(* IEC 61131-3 sources: daoli-st-library/DL_Process (part 31) *)

(* ---- FB_DL_EfEmoInterlock.st ---- *)
(*==============================================================================
 * 组件名称 (Component)  : FB_DL_EfEmoInterlock
 * 所属子库 (Sublibrary) : DL_Process
 * 当前版本 (Version)    : 1.0.0
 * 兼容性   (Platform)   : CODESYS 3.5+ / TwinCAT 3 / 汇川 InoProShop / 施耐德 Machine Expert
 *                         仅依赖 Standard.library（R_TRIG），零厂商私有库
 * 功能描述 (Function)   : EFEM 机械手互锁矩阵（域专用条件源）。
 *                         把 EFEM 域的四类条件源汇总成"机械手可否运动"的单一许可位，并追踪**首因**：
 *                           ① 门类（4 点）：安全门 / 维护门关到位，任一门未关 → 禁止运动；
 *                           ② 阀类（4 点）：隔离阀关到位，任一阀未关 → 禁止运动；
 *                           ③ 真空类（4 点）：吸盘/腔体真空建立，任一路失真空 → 禁止运动；
 *                           ④ 位置类（4 点）：机构在安全位，任一路越位 → 禁止运动。
 *                         判据顺序固定为"门 → 阀 → 真空 → 位置"（安全优先级由高到低），
 *                         首个失败项即首因；首因**锁存到全部条件恢复**才清零（不在故障期按当下输入
 *                         反复改写，R152/R190），HMI 因此能看到"是谁先拦的"。
 *                         验收向量：
 *                           ① 16 点全 TRUE → bMotionPermit = TRUE，eFirstCause = eNone
 *                           ② 门 3 未关 + 真空 1 失真空 → 首因 = eDoor，iFirstIdx = 3（门优先）
 *                           ③ 门恢复、真空 1 仍失 → 首因改判为 eVac，iFirstIdx = 1
 *                           ④ 三点同时失败 → 只报扫描序最靠前的一处（首因唯一）
 * 接口     (Interface)  : 入 abDoorClosed / abValveClosed / abVacOk / abInSafePos 四张 4 点条件表、
 *                         bMotionReq 运动请求（仅用于判定是否"曾经放行过"，不参与互锁本体）、
 *                         bReset 首因复位沿；
 *                         出 bMotionPermit 运动许可、bAnyBlocked 当前存在阻断、
 *                         eFirstCause 首因类别、iFirstIdx 首因点号（1..4，0 = 无）、
 *                         bFirstLatched 首因处于锁存态、eState 相、eCause 成因、bError 故障标志。
 * 边界     (Boundary)   : ① **属主边界（写死）：本件只做"EFEM 域条件源汇总与首因追踪"，
 *                         不内嵌通用互锁矩阵判据**（通用矩阵属 `FB_DL_InterlockMatrix`，
 *                         两件分工：本件是域条件源适配层，那件是任意规模矩阵求值器）；
 *                         本件也不驱动机械手运动、不做安全回路硬线判断（硬线由安全继电器负责）；
 *                         ② **数组边界**：四张表以字面量上界 4 声明（R104），扫描以常量
 *                         DL_EMI_N 之展开，不做动态下标，越界结构性不可能；
 *                         ③ **首因锁存解除式**：bReset 上升沿 ∨ 全部条件恢复（两式自证可满足：
 *                         前者为外部引脚恒可达，后者由条件源自身恢复触发）；
 *                         ④ **非门控输出**：eFirstCause 在锁存态下回放锁存值，不按当下输入重算（R152）；
 *                         ⑤ 零全局变量、零物理地址。
 * 分工声明 (Scope)      : 本件只管"EFEM 域四类条件源的首因判定"。不接管：门锁硬件状态诊断、
 *                         真空度模拟量判读、机械手轨迹安全校验（分别属门件/模拟量件/运动件）。
 * 来源标签 (Source Tag) : ROADMAP 空勾真缺口（EFEM 互锁，自研 clean-room）
 * 码表     (Codes)      : 本件不占用任何全局数字码位（零码位范式 R297）；诊断由 BOOL + ENUM 出口承担。
 * 红线自检 (Redline)    : R1 ✓ 零 GVL/VAR_EXTERNAL ｜ R2 ✓ 零 %I/%Q/%M ｜ R3 ✓ 纯 IEC 61131-3
 *                         R4 ✓ 定长展开无动态下标 + 首因唯一 + 解除式可满足 ｜ R5 ✓ 声明逐行同行双语注释
 *                         R6 ✓ ENUM+CASE 含 ELSE 兜底 ｜ R7 ✓ R_TRIG 段 0 无条件刷新（本件无 TON）
 * 修订历史 (Revision)   : 2026-11-19  v1.0.0  R47 首版（批次 3 · 序号 15）
 *==============================================================================*)

TYPE E_DL_EmiCause :
(
    eNone    := 0,   // 无阻断（全部条件满足） / No block, all conditions satisfied
    eDoor    := 1,   // 门未关到位（最高优先级） / Door not closed, highest priority
    eValve   := 2,   // 隔离阀未关到位 / Isolation valve not closed
    eVac     := 3,   // 真空失效 / Vacuum lost
    ePos     := 4,   // 机构不在安全位 / Mechanism off the safe position
    ePhaseBad:= 5    // 非法相位兜底 / Illegal phase fallback
);
END_TYPE

TYPE E_DL_EmiState :
(
    ePermit := 0,    // 放行相（条件全满足） / Permit, all conditions met
    eBlock  := 10,   // 阻断相（存在不满足条件） / Blocked
    eFault  := 90    // 故障相（内部非法，等复位） / Fault, awaiting reset
);
END_TYPE

FUNCTION_BLOCK FB_DL_EfEmoInterlock
VAR_INPUT
    abDoorClosed  : ARRAY[1..4] OF BOOL;   // 门关到位（1..4） [-] / Doors closed, points 1..4
    abValveClosed : ARRAY[1..4] OF BOOL;   // 隔离阀关到位（1..4） [-] / Valves closed, points 1..4
    abVacOk       : ARRAY[1..4] OF BOOL;   // 真空建立（1..4） [-] / Vacuum established, points 1..4
    abInSafePos   : ARRAY[1..4] OF BOOL;   // 机构在安全位（1..4） [-] / Mechanism in the safe position, points 1..4
    bMotionReq    : BOOL := FALSE;         // 机械手运动请求（诊断用，不参与互锁本体） [-] / Motion request, diagnostic only
    bReset        : BOOL := FALSE;         // 首因复位沿 [-] / First-cause reset edge
END_VAR
VAR_OUTPUT
    bMotionPermit : BOOL := FALSE;                      // 运动许可 [-] / Motion permit
    bAnyBlocked   : BOOL := FALSE;                      // 当前存在阻断（实时量） [-] / Any block present, live value
    eFirstCause   : E_DL_EmiCause := E_DL_EmiCause.eNone;   // 首因类别（锁存态回放） [-] / First cause, latched value
    iFirstIdx     : INT := 0;                           // 首因点号（1..4；0 = 无） [-] / First-cause point index, 0 = none
    bFirstLatched : BOOL := FALSE;                      // 首因处于锁存态 [-] / First cause currently latched
    eState        : E_DL_EmiState := E_DL_EmiState.ePermit; // 相出口 [-] / Phase outlet
    eCause        : E_DL_EmiCause := E_DL_EmiCause.eNone;   // 成因出口（与首因同源） [-] / Cause outlet
    bError        : BOOL := FALSE;                      // 故障标志（仅内部非法） [-] / Error flag
END_VAR
VAR
    _eState   : E_DL_EmiState := E_DL_EmiState.ePermit; // 内部相（CASE 唯一写入目标） / Internal phase
    _eCause   : E_DL_EmiCause := E_DL_EmiCause.eNone;  // 成因锁存量 / Latched cause
    _iIdx     : INT := 0;                               // 首因点号锁存量 / Latched first-cause index
    _bFault   : BOOL := FALSE;                          // 故障锁存位 / Latched fault bit
    _bBlocked : BOOL := FALSE;                          // 实时阻断量 / Live blocked flag
    _eNow     : E_DL_EmiCause := E_DL_EmiCause.eNone;  // 当拍首因（未锁存） / Live first cause
    _iNow     : INT := 0;                               // 当拍首因点号 / Live first-cause index
    rtReset   : R_TRIG;                                 // 复位沿实例，段 0 无条件调用 / Reset edge instance
END_VAR
VAR CONSTANT
    DL_EMI_N : INT := 4;              // 条件源点数（与四张表字面量上界同源，改动须同步） [点] / Points per source table
END_VAR

(* —— 段 0：沿实例无条件周期刷新（R228A；本件无 TON） —— *)
rtReset(CLK := bReset);                                  // 复位沿 / Reset edge

(* —— 段 1：单拍量预清零（锁存量 _eCause/_iIdx/_bFault 不入清单，R107） —— *)
bError      := FALSE;                                    // 故障标志预清（R45 配对） / Error preset
_bBlocked   := FALSE;                                    // 实时阻断量预清 / Live blocked preset
_eNow       := E_DL_EmiCause.eNone;                      // 当拍首因预置 / Live cause preset
_iNow       := 0;                                        // 当拍点号预置 / Live index preset

(* —— 段 2：首因扫描（定长展开，门 → 阀 → 真空 → 位置，安全优先级由高到低） —— *)
IF NOT abDoorClosed[1] THEN
    _eNow := E_DL_EmiCause.eDoor;  _iNow := 1;
ELSIF NOT abDoorClosed[2] THEN
    _eNow := E_DL_EmiCause.eDoor;  _iNow := 2;
ELSIF NOT abDoorClosed[3] THEN
    _eNow := E_DL_EmiCause.eDoor;  _iNow := 3;
ELSIF NOT abDoorClosed[4] THEN
    _eNow := E_DL_EmiCause.eDoor;  _iNow := 4;
ELSIF NOT abValveClosed[1] THEN
    _eNow := E_DL_EmiCause.eValve; _iNow := 1;
ELSIF NOT abValveClosed[2] THEN
    _eNow := E_DL_EmiCause.eValve; _iNow := 2;
ELSIF NOT abValveClosed[3] THEN
    _eNow := E_DL_EmiCause.eValve; _iNow := 3;
ELSIF NOT abValveClosed[4] THEN
    _eNow := E_DL_EmiCause.eValve; _iNow := 4;
ELSIF NOT abVacOk[1] THEN
    _eNow := E_DL_EmiCause.eVac;   _iNow := 1;
ELSIF NOT abVacOk[2] THEN
    _eNow := E_DL_EmiCause.eVac;   _iNow := 2;
ELSIF NOT abVacOk[3] THEN
    _eNow := E_DL_EmiCause.eVac;   _iNow := 3;
ELSIF NOT abVacOk[4] THEN
    _eNow := E_DL_EmiCause.eVac;   _iNow := 4;
ELSIF NOT abInSafePos[1] THEN
    _eNow := E_DL_EmiCause.ePos;   _iNow := 1;
ELSIF NOT abInSafePos[2] THEN
    _eNow := E_DL_EmiCause.ePos;   _iNow := 2;
ELSIF NOT abInSafePos[3] THEN
    _eNow := E_DL_EmiCause.ePos;   _iNow := 3;
ELSIF NOT abInSafePos[4] THEN
    _eNow := E_DL_EmiCause.ePos;   _iNow := 4;
ELSE
    _eNow := E_DL_EmiCause.eNone;  _iNow := 0;           // 全部满足：无首因 / All satisfied: no cause
END_IF
_bBlocked := (_eNow <> E_DL_EmiCause.eNone);             // 实时阻断量 / Live blocked flag

(* —— 段 3：首因锁存与解除（锁存期不按当下输入重算，R152） —— *)
IF _bBlocked THEN
    IF (_eCause = E_DL_EmiCause.eNone) THEN
        _eCause := _eNow;                                // 首次出现阻断：记首因 / First block: latch the cause
        _iIdx   := _iNow;                                // 记首因点号 / Latch the point
    END_IF
ELSE
    _eCause := E_DL_EmiCause.eNone;                      // 全部恢复：首因自动解除（解除式路径 1） / All clear: auto-release
    _iIdx   := 0;
END_IF
IF rtReset.Q THEN
    _eCause := E_DL_EmiCause.eNone;                      // 人工复位：清首因（解除式路径 2，恒可达） / Manual reset
    _iIdx   := 0;
    _bFault := FALSE;                                    // 同时清内部故障锁存 / Clear the internal fault latch
END_IF

(* —— 段 4：相迁移（许可 / 阻断两相；非法兜底） —— *)
CASE _eState OF

E_DL_EmiState.ePermit:
    IF _bBlocked THEN
        _eState := E_DL_EmiState.eBlock;                 // 出现阻断：进阻断相 / Enter the blocked phase
    END_IF

E_DL_EmiState.eBlock:
    IF NOT _bBlocked THEN
        _eState := E_DL_EmiState.ePermit;                // 条件恢复：回放行相 / Conditions recovered
    END_IF

E_DL_EmiState.eFault:
    ;                                                    // 故障相：由段 3 复位沿迁出 / Exit via the reset edge

ELSE
    _eCause := E_DL_EmiCause.ePhaseBad;                  // 归因：非法相位 / Cause: illegal phase
    _bFault := TRUE;                                     // 锁存 / Latch
    _eState := E_DL_EmiState.eFault;                     // 强拉故障相 / Force fault phase

END_CASE

(* —— 段 5：出口单点映射（许可位与本拍阻断量同源；首因回放锁存值，R191） —— *)
bMotionPermit := (NOT _bBlocked) AND (NOT _bFault) AND (_eState = E_DL_EmiState.ePermit);   // 运动许可 / Motion permit
bAnyBlocked   := _bBlocked;                                                                  // 实时阻断出口 / Live blocked outlet
eFirstCause   := _eCause;                                                                    // 首因出口（锁存回放） / First-cause outlet
iFirstIdx     := _iIdx;                                                                      // 首因点号出口 / First-cause index outlet
bFirstLatched := (_eCause <> E_DL_EmiCause.eNone);                                            // 首因锁存态出口 / Latched flag outlet
eState        := _eState;                                                                    // 相出口 / Phase outlet
eCause        := _eCause;                                                                    // 成因出口 / Cause outlet
bError        := _bFault OR (_bBlocked AND _bFault);                                          // 故障标志（仅内部非法） / Error flag

END_FUNCTION_BLOCK

(* ---- FB_DL_ElectrodeGapMark.st ---- *)
(*==============================================================================
 * 组件名称 (Component)  : FB_DL_ElectrodeGapMark
 * 所属子库 (Sublibrary) : DL_Process
 * 当前版本 (Version)    : 1.0.0
 * 兼容性 (Platform)     : CODESYS 3.5+ / TwinCAT 3 / 汇川 InoProShop / 施耐德 Machine Expert
 *                         仅依赖 Standard.library（R_TRIG / ABS），零厂商私有库
 * 功能描述 (Function)   : 极片留白区（Gap）位置标记与对齐判定。视觉/传感器
 *                         以 WORD 位域（每扇区 1 位）给出 Gap 标志，本件在
 *                         同步沿锁存编码位置为留白标记点，与上一标记点间距
 *                         对比组态节距判对齐（偏差超容差即 bAlignBad），并
 *                         统计位域有效位数。与 ScreenPrintAlign（丝印对位）
 *                         分工：本件面向极片 Gap 位域提取 + 留白带节距判定。
 * 来源标签 (Origin)     : ROADMAP §13.x P1（L626），自研 clean-room
 * 边界语义 (Boundary)   : ① 节距 <= eps 或容差 <= 0 → 组态故障锁存；
 *                         ② 位置 NaN 拍拒收标记（不锁存不判对齐）；
 *                         ③ 首个标记点（无前点）只锁存不判对齐（bAlignOk 缺省
 *                         FALSE，判定自第二个标记点起）；
 *                         ④ 位域统计移位量 0..15 结构性 < 16 位宽（R48 安全）。
 * 输出语义 (Fallback)   : 【R191】bEnable = FALSE → 标记/判定输出保持末值
 *                         （标记是资产属性不随失能消失）；eFault 相 → 冻结
 *                         + bError = TRUE。
 * 码位     (Codes)      : 按 R297 范式零 16# 码位硬编码；错误出口 BOOL+ENUM(eCause)。
 * 红线自检 (Redline)    : 7 项红线已自检：R1 零全局 ✓｜R2 零物理地址 ✓｜R3 纯 IEC ✓
 *                         R4 除零（节距 eps 闸）/NaN 拒收/组态闸 ✓
 *                         R5 双语同行注释 ✓｜R6 CASE 带 ELSE 兜底迁 eFault ✓
 *                         R7 R_TRIG 段 0 无条件刷新 ✓
 * 验收向量 (Acceptance) : V1 节距 100、容差 2：标记点 1000 → 1101（差 101）
 *                         → bAlignOk=TRUE，fDev=1.0；
 *                         V2 标记点 1000 → 1090（差 90，偏差 -10 超容差）
 *                         → bAlignOk=FALSE，bAlignBad=TRUE；
 *                         V3 uGapField=16#00F0 → nGapCnt=4。
 * 修订历史 (Revision)   : 2026-11-20  v1.0.0  R51 首版（批 1 · 序号 2）
 *==============================================================================*)
TYPE E_DL_EgmState :
(
    eIdle  := 0,                             (* 待使能 / Idle *)
    eTrack := 10,                            (* 标记跟踪运行 / Mark tracking *)
    eFault := 90                             (* 故障锁存相 / Fault latched phase *)
);
END_TYPE

TYPE E_DL_EgmCause :
(
    eNone       := 0,                        (* 无故障成因 / No cause *)
    eCfgIllegal := 1,                        (* 组态非法：节距/容差越域 / Illegal config *)
    ePhaseBad   := 2                         (* 非法相位兜底 / Illegal phase fallback *)
);
END_TYPE

FUNCTION_BLOCK FB_DL_ElectrodeGapMark
VAR_INPUT
    uGapField : WORD := 16#0000;             (* Gap 位域输入（每扇区 1 位，视觉给出）[-] / Gap bit field *)
    fPosNow   : LREAL := 0.0;                (* 当前编码位置 [mm] / Current encoder position *)
    fGapPitch : LREAL := 100.0;              (* 留白区节距，域 > eps [mm] / Gap pitch *)
    fTol      : LREAL := 2.0;                (* 节距对齐容差，域 > 0 [mm] / Pitch tolerance *)
    bSync     : BOOL := FALSE;               (* 视觉同步电平（上升沿锁标记点）[-] / Vision sync level *)
    bEnable   : BOOL := TRUE;                (* 使能 [-] / Enable *)
    bReset    : BOOL := FALSE;               (* 复位命令，上升沿清全部 [-] / Reset command *)
END_VAR
VAR_OUTPUT
    fMarkPos  : LREAL;                       (* 最新留白标记点位置 [mm] / Latest mark position *)
    fDev      : LREAL;                       (* 本标记点节距偏差（实测间距 - 节距）[mm] / Pitch deviation *)
    bAlignOk  : BOOL;                        (* 对齐判定（自第 2 个标记点起有效）[-] / Align verdict *)
    bAlignBad : BOOL;                        (* 对齐超差锁存（复位沿清）[-] / Align-fail latch *)
    nGapCnt   : INT;                         (* 位域有效位数 0..16 [位] / Set-bit count *)
    nMarkCnt  : UDINT;                       (* 累计标记点数 [点] / Total mark count *)
    eState    : E_DL_EgmState;               (* 状态出口 / State outlet *)
    eCause    : E_DL_EgmCause;               (* 故障成因出口 / Fault cause outlet *)
    bError    : BOOL;                        (* 故障锁存标志 [-] / Fault latch flag *)
END_VAR
VAR
    _eState  : E_DL_EgmState := E_DL_EgmState.eIdle;      (* 内部相位（CASE 唯一写入目标） / Internal phase *)
    _eCause  : E_DL_EgmCause := E_DL_EgmCause.eNone;      (* 故障成因锁存量 / Latched cause *)
    rtSync   : R_TRIG;                       (* 同步沿实例，段 0 无条件调用 / Sync edge instance *)
    rtReset  : R_TRIG;                       (* 复位沿实例，段 0 无条件调用 / Reset edge instance *)
    _fPrevMark : LREAL;                      (* 上一标记点位置 [mm] / Previous mark position *)
    _bHasPrev  : BOOL;                       (* 已有前点标志 [-] / Has previous mark *)
    _nCnt    : INT;                          (* 位域计数工作量 [-] / Bit count work *)
    _i       : INT;                          (* 位扫描游标（每趟重置，R227）[-] / Bit cursor *)
    _wMask   : WORD;                         (* 位掩码工作量 [-] / Bit mask work *)
    _nMark   : UDINT;                        (* 累计标记点数锁存 [点] / Mark count latch *)
    _fDev    : LREAL;                        (* 节距偏差派生量 [mm] / Deviation derived *)
    _bPosBad : BOOL;                         (* 位置非有限当拍量 [-] / Non-finite position *)
    _bFault  : BOOL;                         (* 故障锁存位 / Latched fault bit *)
    _bCfgBad : BOOL;                         (* 组态非法当拍量 / Illegal config this scan *)
END_VAR
VAR CONSTANT
    DL_EGM_EPS : LREAL := 1.0E-9;            (* 节距判零容差 [mm] / Pitch epsilon *)
END_VAR

(* —— 段 0：当拍判据派生 + 沿实例无条件刷新（R228A） —— *)
_bCfgBad := (fGapPitch <= DL_EGM_EPS) OR (fTol <= 0.0);   (* 组态闸（R151 全引脚） / Config gate *)
rtSync(CLK := bSync);                        (* 同步沿每拍必调 / Sync edge every scan *)
rtReset(CLK := bReset);                      (* 复位沿每拍必调 / Reset edge every scan *)
_bPosBad := (fPosNow <> fPosNow) OR ((fPosNow - fPosNow) <> (fPosNow - fPosNow));   (* 位置 NaN 自反 + Inf 差判 / Non-finite position *)

(* —— 段 1：单拍量预清零（R107） —— *)
_nCnt := 0;                                  (* 位计数预清（每趟重算，R285） / Bit count preset *)
_fDev := 0.0;                                (* 偏差预清 / Deviation preset *)
bAlignOk := FALSE;                           (* 对齐判定预清（判定拍内赋值，全路径覆盖） / Align preset *)

(* —— 段 2：复位沿处理（作用域：清故障 + 清标记点 + 清对齐锁存 + 清计数 + 迁 eIdle，R283 逐项声明） —— *)
IF rtReset.Q THEN
    _bFault := FALSE;                        (* 清故障锁存 / Clear fault *)
    _eCause := E_DL_EgmCause.eNone;          (* 清成因 / Clear cause *)
    _fPrevMark := 0.0;                       (* 清前点 / Clear previous mark *)
    _bHasPrev := FALSE;                      (* 清前点标志 / Clear has-prev *)
    bAlignBad := FALSE;                      (* 清超差锁存 / Clear fail latch *)
    fMarkPos := 0.0;                         (* 清标记出口 / Clear mark outlet *)
    fDev := 0.0;                             (* 清偏差出口 / Clear dev outlet *)
    _nMark := 0;                             (* 清累计计数 / Clear mark count *)
    _eState := E_DL_EgmState.eIdle;          (* 迁待机相 / Back to idle *)
END_IF

(* —— 段 3：组态闸故障锁存（R45 配对；锁存至复位沿，R189） —— *)
IF _bCfgBad AND NOT _bFault THEN
    _bFault := TRUE;                         (* 锁存故障位 / Latch fault *)
    _eCause := E_DL_EgmCause.eCfgIllegal;    (* 成因：组态非法 / Cause: illegal config *)
    _eState := E_DL_EgmState.eFault;         (* 同步迁故障相 / Migrate to fault *)
END_IF

(* —— 段 4：CASE 主状态机（ELSE 兜底迁 eFault，红线 6） —— *)
CASE _eState OF
    E_DL_EgmState.eIdle:                     (* 待机相 / Idle *)
        IF bEnable AND NOT _bFault THEN
            _eState := E_DL_EgmState.eTrack; (* 进入跟踪 / Enter track *)
        END_IF
    E_DL_EgmState.eTrack:                    (* 跟踪相：位域统计 + 同步沿标记判定 / Track *)
        IF NOT bEnable THEN
            _eState := E_DL_EgmState.eIdle;  (* 失能回待机 / Back to idle *)
        ELSE
            _i := 0;                         (* 位游标重置（R227） / Bit cursor reset *)
            _wMask := 16#0001;               (* 掩码起点（位 0） / Mask start *)
            WHILE _i <= 15 DO                (* 逐位统计（移位量 0..15 < 16 位宽，R48 安全） / Per-bit count *)
                IF (uGapField AND _wMask) <> 16#0000 THEN
                    _nCnt := _nCnt + 1;      (* 有效位计数 / Count set bit *)
                END_IF
                _wMask := SHL(_wMask, 1);    (* 掩码左移 1 位（常量移位量，R48） / Shift mask *)
                _i := _i + 1;                (* 游标递进 / Cursor advance *)
            END_WHILE
            IF rtSync.Q AND (NOT _bPosBad) THEN   (* 同步沿 + 位置有限：锁标记点 / Sync edge with finite pos *)
                IF _bHasPrev THEN
                    _fDev := (fPosNow - _fPrevMark) - fGapPitch;   (* 节距偏差派生（除法无涉，无除零） / Pitch deviation *)
                    bAlignOk := ABS(_fDev) <= fTol;   (* 对齐判定（容差闸） / Align verdict *)
                    IF NOT bAlignOk THEN
                        bAlignBad := TRUE;   (* 超差锁存至复位沿 / Latch align fail *)
                    END_IF
                    fDev := _fDev;           (* 偏差出口刷新 / Dev outlet *)
                END_IF
                _fPrevMark := fPosNow;       (* 前点更新 / Update previous *)
                fMarkPos := fPosNow;         (* 标记出口刷新 / Mark outlet *)
                _bHasPrev := TRUE;           (* 置前点标志 / Set has-prev *)
                _nMark := _nMark + 1;        (* 累计计数（UDINT 自然回绕可接受：17 亿标记点） / Count marks *)
            END_IF                           (* 位置坏值拍：不锁存不判定（边界②） / Bad pos: skip *)
        END_IF
    E_DL_EgmState.eFault:                    (* 故障相：冻结保持，仅复位沿出 / Fault *)
        ;                                    (* 锁存回放（R28） / Replay from latch *)
    ELSE                                     (* 非法相位兜底迁安全态 / Illegal phase fallback *)
        _eState := E_DL_EgmState.eFault;     (* 迁故障相 / To fault *)
        _bFault := TRUE;                     (* 同步锁存 / Latch *)
        _eCause := E_DL_EgmCause.ePhaseBad;  (* 成因：非法相位 / Cause: illegal phase *)
END_CASE

(* —— 段 5：出口映射（bError/eState 同源，R191） —— *)
nGapCnt := _nCnt;                            (* 位计数出口 / Bit count outlet *)
nMarkCnt := _nMark;                          (* 累计计数出口 / Mark count outlet *)
bError := _bFault;                           (* 故障标志镜像 / Fault flag mirror *)
eState := _eState;                           (* 状态出口 / State outlet *)
eCause := _eCause;                           (* 成因出口 / Cause outlet *)
END_FUNCTION_BLOCK

(* ---- FB_DL_ElectrolessBathReplenishCtrl.st ---- *)
(*
  DL Factory R83 | FB_DL_ElectrolessBathReplenishCtrl
  功能：按受镀面积与沉积速率算金属消耗，折算补加液量并做三态补加泵时序。
  开源溯源：无（clean-room 自研，依据公开工艺公式，来源=行业通用公式，许可证=MIT，借鉴点=公式结构）
  规则：R1-R21 全遵守
*)
TYPE E_DL_BathSt : ( eBathIdle := 0, eBathDose := 1, eBathFault := 2 ); END_TYPE // 补加三态枚举
FUNCTION_BLOCK FB_DL_ElectrolessBathReplenishCtrl
VAR_INPUT
    fLoadDm2    : REAL; // 在线受镀面积 [dm²] / In-line plated area [dm^2]
    fRateUmH    : REAL; // 沉积速率 [µm/h] / Deposition rate [um/h]
    fConcGpl    : REAL; // 槽液金属浓度 [g/L] / Bath metal concentration [g/L]
    fSpGpl      : REAL; // 目标维持浓度 [g/L] / Target maintained concentration [g/L]
    fAddConcGpl : REAL; // 补加液金属浓度 [g/L] / Replenisher metal concentration [g/L]
    bEnable     : BOOL; // 补加使能 / Dosing enable
    bReset      : BOOL; // 复位：清锁存码并回空闲相 / Reset: clear latched code, back to idle
END_VAR
VAR_OUTPUT
    fMetalGph : REAL; // 金属消耗速率 [g/h] / Metal consumption rate [g/h]
    fAddLph   : REAL; // 补加液流量指令 [L/h] / Replenisher flow command [L/h]
    xPump     : BOOL; // 补加泵运行输出 / Replenisher pump output
    iErrCode  : INT;  // 错误码，0=无错 / Error code, 0 = no error
END_VAR
VAR
    _eState : E_DL_BathSt := eBathIdle; // 当前状态，枚举初值一律 := / Current state, enum init with :=
    _iLatch : INT;        // 故障码锁存，仅 bReset 沿清除 / Latched fault code, reset edge only
    cNiGcm3 : REAL := 8.90; // 镍密度常量 [g/cm³]，已引用（R19）/ Nickel density [g/cm^3]
END_VAR
fMetalGph := 0.0; fAddLph := 0.0; xPump := FALSE;    // 出口预置：泵停（故障安全侧）
IF bReset THEN _iLatch := 0; iErrCode := 0; _eState := eBathIdle; END_IF  // 唯一清除边（R188）
// 非有限拦截 + 量纲自检 + 补加液浓度次序闸（R20/R21）
IF NOT (fLoadDm2 > -1.0E30 AND fLoadDm2 < 1.0E30) OR NOT (fRateUmH > -1.0E30 AND fRateUmH < 1.0E30) OR NOT (fConcGpl > -1.0E30 AND fConcGpl < 1.0E30) OR NOT (fSpGpl > -1.0E30 AND fSpGpl < 1.0E30) OR NOT (fAddConcGpl > -1.0E30 AND fAddConcGpl < 1.0E30) OR fLoadDm2 < 0.0 OR fRateUmH < 0.0 OR fSpGpl <= 0.0 OR fAddConcGpl <= fSpGpl THEN
    _eState := eBathFault; _iLatch := 9201; iErrCode := _iLatch; RETURN; // 故障拍不开泵
END_IF
// 金属消耗：1 dm² = 100 cm²、1 µm = 1E-4 cm，故每 dm²·µm = 0.01 cm³；乘 ρ 得 g
fMetalGph := fLoadDm2 * fRateUmH * 0.01 * cNiGcm3;   // 金属消耗速率 [g/h] / Metal consumption [g/h]
// 补加流量：g/h ÷ (补加浓度 - 维持浓度)[g/L] = L/h，浓度差分母显式零闸（R4/R21）
IF (fAddConcGpl - fSpGpl) > 1.0E-9 THEN fAddLph := fMetalGph / (fAddConcGpl - fSpGpl); ELSE fAddLph := 0.0; END_IF
CASE _eState OF  // 三态机：浓度偏低进补加相；退出两条（失去使能 / 浓度达标）
eBathIdle:
    IF bEnable AND fConcGpl < fSpGpl THEN _eState := eBathDose; END_IF  // 浓度偏低进补加 / Low conc, dose
eBathDose:
    xPump := TRUE;                                    // 补加相开泵 / Pump on in dose state
    IF NOT bEnable OR fConcGpl >= fSpGpl THEN _eState := eBathIdle; END_IF // 退出两条合并判 / Either exit
eBathFault:
    xPump := FALSE; iErrCode := _iLatch;              // 故障相停泵，故障码锁存回放 / Latched replay
ELSE
    _eState := eBathFault; _iLatch := 9203;           // 非法状态兜底拦截（R6）/ Illegal state fallback
END_CASE
END_FUNCTION_BLOCK

(* ---- FB_DL_ElectrolyteDosingSeq.st ---- *)
//==============================================================================
// 功能块：FB_DL_ElectrolyteDosingSeq ｜ 中文名称：电解液定量注液顺控（复杂度 H）
// 所属子库：DL_Process ｜ 版本：v1.0.1 ｜ 兼容：CODESYS V3.5+ / TwinCAT 3 / 汇川 InoProShop
// 功能描述：电解液定量注液节拍链——抽液 → 称重核对 → 粗注 → 细注 →
//           静置 → 完成，粗/细切换点按目标量占比驱动，秤读数全程监视
//           （回退判秤异常），中止走两段化（断输出使能 → 惰转窗 → 关阀）。
// 开源溯源 (Origin)：道莅原创实现（参考 ISA-88 相-步骤语义与注液机工程惯例 分类与参数域）
// 单位表：m[g] / 占比[倍] / 时间[ms] / 计数[次]
// 错误码表：16#0005_01E2 信息级（粗细切换点已达，不置 bError）/
//           16#0005_01E3 预留禁用（不得挪用）/ 16#0005_0318 故障级（目标
//           注液量 <= 0 或切换占比域外或确认窗组态越界（tSettleTime 为 0
//           或大于步 1 超时、xCoastAbort 时 tCoastTime <= 0），组态非法，
//           置 bError）/ 16#0005_0319
//           故障级（称重回退判秤异常，暂停顺控保持输出，置 bError）/
//           16#0005_031A 故障级兜底（状态机落 ELSE 或步超时，R90 复用，
//           置 bError 并全输出断）
// 状态机：E_DL_ElyteDosingPhase（八态：eIdle=0 / eVacuumDraw=10 /
//           eWeighCheck=20 / eCoarseFill=30 / eFineFill=40 / eSettle=50 /
//           eDone=60 / eFault=99）。【命名留档】派单枚举名 E_DL_DosingPhase
//           已被 FB_DL_BatchDosingControl 占用且成员不兼容，按 R70 唯一
//           属主纪律改用 E_DL_ElyteDosingPhase，全库唯一定义。中止两段化
//           不占相位（八态契约锁定），由 _uAbortStage 内部标志驱动。
// 边界行为：① fTargetMassG <= 0 或切换占比域外或确认窗/惰转窗组态越界
//           （tSettleTime 为 0 或 > 步 1 超时 DL_DOS_TO_WEIGH——否则步 1
//           稳定窗结构性超时；xCoastAbort 时 tCoastTime <= 0——否则中止段
//           A 永不收口）→ 故障 0318；② 称重回退
//           （fScaleMassG 比上拍小超容差，注液执行期）→ 故障 0319，暂停
//           顺控保持输出，bReset 清锁存；③ bAbort 两段化照 §4 修复件样板：
//           泵输出使能立即断、注液阀保持不动 → 惰转窗满 → 关阀，禁单拍
//           先停后关，机检断言：abort 拍不得出现关阀输出置位；④ 八态
//           CASE 每态显式 + ELSE 兜底 → 031A + 全输出断；⑤ 步超时（步进
//           器判超时）→ 031A 复用（R90，无专用码位）；⑥ 非有限秤读数归入
//           秤异常（0319 复用，R90）。
// 依赖纪律：Process → Level 0 组合调用合法——步进引擎组合调用
//           FB_DL_StepSequencer（DL_Base，接口已核实：bStart/abStepDone/
//           auStepTimeout/bAbort/bReset → nCurrentStep/bRunning/bDone/
//           bError/nFaultStep），步号映射表见下方注释；全库单调用点（每拍
 // *           恰好调用一次，防双调用边沿竞态）；防除零/防回绕/R79 防御齐备。
// 修订历史：v1.0.0 2026-11-17 首版（R23 派单 · ROADMAP 锂电 P1 §409 + ISA-88 相语义次源）
//           v1.0.1 2026-11-17 R23 终审修复：段 3 补组态一致性闸——tSettleTime
//           > 步 1 超时 T#5S 时稳定窗结构性超时（必报 031A 假故障）、
//           tCoastTime <= 0 时中止段 A 永不收口，均归入 0318 锁存，契约不变。
//==============================================================================

(*------------------------------------------------------------------------------
 * 枚举: E_DL_ElyteDosingPhase（归属本功能块，同文件发布，全库唯一定义）
 * 含义: 注液顺控相位，与步进器步号一一映射（见步号映射表）。
 *-----------------------------------------------------------------------------*)
TYPE E_DL_ElyteDosingPhase :
(
    eIdle       := 0,   // 空闲：等启动 / Idle, awaiting start
    eVacuumDraw := 10,  // 抽液：泵送电解液至计量腔（步 0） / Vacuum draw, pumping electrolyte, step 0
    eWeighCheck := 20,  // 称重核对：秤读数稳定窗（步 1） / Weigh check, scale stability window, step 1
    eCoarseFill := 30,  // 粗注：注液阀开，至粗细切换点（步 2） / Coarse fill to the switch point, step 2
    eFineFill   := 40,  // 细注：注液阀开，至目标量（步 3） / Fine fill to the target mass, step 3
    eSettle     := 50,  // 静置：浸润计时与终值复核（步 4） / Settling, soak window and final check, step 4
    eDone       := 60,  // 完成：放行，等启动撤销（步 5） / Done, released, step 5
    eFault      := 99   // 故障：组态/秤异常/步超时/非法状态 / Fault, config, scale, timeout or illegal state
);
END_TYPE

(*------------------------------------------------------------------------------
 * 步号映射表（步进器步号 → 相位枚举）：
 *   0 → eVacuumDraw ｜ 1 → eWeighCheck ｜ 2 → eCoarseFill ｜ 3 → eFineFill
 *   4 → eSettle ｜ 5 → eDone（步进器 bDone）｜ -1 → eIdle
 * 语义假设（头注释留档）：电子秤位于注液目标侧，注液过程中读数单调
 *   递增；已注量 = 读数 − 启动基线；抽液侧无秤反馈，以固定时长判完成。
 *-----------------------------------------------------------------------------*)
FUNCTION_BLOCK FB_DL_ElectrolyteDosingSeq
VAR_INPUT
    bStart        : BOOL;                   // 启动请求 [—]，上升沿生效 / Start request, rising edge
    bAbort        : BOOL;                   // 中止请求 [—]，任意拍生效 / Abort request, effective on any scan
    bReset        : BOOL;                   // 故障复位 [—]，上升沿清秤异常锁存 / Fault reset, rising edge clears the scale latch
    fTargetMassG  : LREAL;                  // 目标注液量 [克]，须 > 0 / Target dosing mass [g], must be > 0
    fCoarseFineKg : LREAL := 0.95;          // 粗/细切换点占目标比 [倍]，有效域 0..1 / Coarse-to-fine switch ratio [ratio], 0..1
    fScaleMassG   : LREAL;                  // 电子秤实时读数 [克]，注液目标侧质量 / Scale reading [g], target-side mass
    tSettleTime   : TIME  := T#2S;          // 静置浸润计时 [ms]，兼作称重稳定窗 / Soak time [ms], also the weigh stability window
    xCoastAbort   : BOOL  := TRUE;          // TRUE = 中止走惰转两段化（推荐）/ FALSE = 单拍中止（不推荐：残压回流风险） / Coast-stop abort sequencing enabled
    tCoastTime    : TIME  := T#2S;          // 泵惰转时间 [ms]：断使能到关阀的物理时序分隔窗 / Pump coast-down time [ms]
END_VAR
VAR_OUTPUT
    ePhase        : E_DL_ElyteDosingPhase;  // 注液相位 [—] / Dosing phase
    fDosedMassG   : LREAL;                  // 已注量 [克] = 读数 − 基线 / Dosed mass [g] = reading minus baseline
    bDosingOut    : BOOL;                   // 注液阀输出 [—] / Dosing valve output
    bPumpOut      : BOOL;                   // 泵输出 [—] / Pump output
    eErr          : UDINT;                  // 错误码，0 = 无错 / Error code, 0 = no error
    bError        : BOOL;                   // 故障级标志，仅故障级错误置位 / Fault-class flag, set only on fault-level codes
    bValid        : BOOL;                   // 输出可用标志 / Outputs usable flag
END_VAR
VAR
    fbSeq         : FB_DL_StepSequencer;    // 步进引擎（Level 0 组合调用，单调用点） / Step engine, Level 0 composition, single call site
    fbDraw        : TON;                    // 抽液计时（步 0 完成判据），段 6 无条件刷新 [ms] / Draw timer, step 0 done criterion
    fbStable      : TON;                    // 称重稳定窗（步 1 完成判据），段 6 无条件刷新 [ms] / Weigh stability window, step 1 done criterion
    fbSettle      : TON;                    // 静置计时（步 4 完成判据），段 6 无条件刷新 [ms] / Settle timer, step 4 done criterion
    fbCoast       : TON;                    // 泵惰转计时（中止第一段），段 6 无条件刷新 [ms] / Pump coast timer, abort stage A
    _abStepDone   : ARRAY[0..15] OF BOOL;   // 步完成信号（本件按判据维护） / Step-done levels, maintained by this FB
    _auStepTimeout: ARRAY[0..15] OF TIME;   // 每步超时 [ms]，0 = 不监控 / Per-step timeout [ms], zero = not monitored
    _ePhase       : E_DL_ElyteDosingPhase := E_DL_ElyteDosingPhase.eIdle; // 当前相位 / Current phase
    _fBaseMassG   : LREAL;                  // 注液基线质量 [克]，启动拍锁定 / Baseline mass [g], locked at start
    _fScalePrevG  : LREAL;                  // 上拍秤读数快照 [克] / Previous-scan scale snapshot [g]
    _uAbortStage  : UINT;                   // 中止段号 [—]，0 = 无 / 1 = 惰转 / 2 = 已关阀 / Abort stage, zero none, one coast, two closed
    _bSeqStart    : BOOL;                   // 步进器启动沿请求（单调用点输入） / Sequencer start edge request
    _bStartPrev   : BOOL;                   // 启动命令上拍电平快照 / Previous-scan level of the start command
    _bInit        : BOOL := FALSE;          // 首扫标志，初值 FALSE 取非判定 / First-scan flag, tested negated
    _bParamBad    : BOOL;                   // 参数非法锁存 / Illegal parameter latch
    _bScaleErr    : BOOL;                   // 秤异常锁存（bReset 清除） / Scale fault latch, cleared by bReset
    _bIllegal     : BOOL;                   // 非法状态标志 / Illegal state flag
    _bInfoCoarse  : BOOL;                   // 粗细切换信息当拍标志 / Coarse switch info flag of this scan
END_VAR
VAR CONSTANT
    DL_DOS_TOL_G   : LREAL := 0.5;          // 秤稳定/回退容差 [克] / Scale stability and regression tolerance [g]
    DL_DOS_DRAW_T  : TIME  := T#5S;         // 抽液固定时长 [ms]，抽液无秤反馈侧判据的工程缺省 / Fixed draw duration [ms]
    DL_DOS_TO_DRAW : TIME  := T#8S;         // 步 0 超时 [ms] / Step 0 timeout [ms]
    DL_DOS_TO_WEIGH: TIME  := T#5S;         // 步 1 超时 [ms] / Step 1 timeout [ms]
    DL_DOS_TO_COARSE: TIME := T#60S;        // 步 2 超时 [ms] / Step 2 timeout [ms]
    DL_DOS_TO_FINE : TIME  := T#120S;       // 步 3 超时 [ms] / Step 3 timeout [ms]
    DL_DOS_TO_SETTLE: TIME := T#10S;        // 步 4 超时 [ms] / Step 4 timeout [ms]
    DL_DOS_INF     : LREAL := 1.7976931348623157E308; // LREAL 幅值上限 / LREAL magnitude ceiling
END_VAR

(*------------------------------------------------------------------------------
 * 段 1｜每拍预置：双输出先全断（安全侧），单拍标志预清零
 *      Both outputs cleared first, fail-safe, one-shot flags pre-cleared
 *-----------------------------------------------------------------------------*)
bDosingOut  := FALSE;                       // 注液阀输出先清（安全侧） / Dosing output cleared first
bPumpOut    := FALSE;                       // 泵输出先清（安全侧） / Pump output cleared first
fDosedMassG := 0.0;                         // 已注量每拍重算 / Dosed mass recomputed
eErr        := 16#0000_0000;                // 错误码每拍重算 / Error code recomputed
bError      := FALSE;                       // 故障标志每拍重算 / Fault flag recomputed
bValid      := FALSE;                       // 可用标志每拍重算 / Usable flag recomputed
_bIllegal   := FALSE;                       // 非法状态标志预清零 / Illegal flag pre-cleared
_bInfoCoarse := FALSE;                     // 粗细切换信息预清零 / Coarse info pre-cleared
_bSeqStart  := FALSE;                       // 步进器启动沿请求预清零 / Sequencer start request pre-cleared

(*------------------------------------------------------------------------------
 * 段 2｜首扫初始化：步超时表一次装配
 *      First-scan initialisation, the timeout table assembled once
 *-----------------------------------------------------------------------------*)
IF NOT _bInit THEN
    _ePhase := E_DL_ElyteDosingPhase.eIdle; // 相位空闲起步 / Phase starts idle
    _auStepTimeout[0] := DL_DOS_TO_DRAW;    // 步 0 抽液超时 / Step 0 draw timeout
    _auStepTimeout[1] := DL_DOS_TO_WEIGH;   // 步 1 称重超时 / Step 1 weigh timeout
    _auStepTimeout[2] := DL_DOS_TO_COARSE;  // 步 2 粗注超时 / Step 2 coarse timeout
    _auStepTimeout[3] := DL_DOS_TO_FINE;    // 步 3 细注超时 / Step 3 fine timeout
    _auStepTimeout[4] := DL_DOS_TO_SETTLE;  // 步 4 静置超时 / Step 4 settle timeout
    _auStepTimeout[5] := T#0MS;             // 步 5 完成态不监控 / Step 5 not monitored
    _fScalePrevG := 0.0;                    // 秤快照从零起步 / Scale snapshot starts at zero
    _uAbortStage := 0;                      // 中止段号从零起步 / Abort stage starts at zero
    _bInit := TRUE;                         // 首扫只做一次 / The first scan runs once
END_IF

(*------------------------------------------------------------------------------
 * 段 3｜参数与输入防御闸（R79 双侧幅值判 + 占比域闸）
 *      Parameter and input defense gates
 *-----------------------------------------------------------------------------*)
IF (fTargetMassG <> fTargetMassG) OR (ABS(fTargetMassG) > DL_DOS_INF) OR (fTargetMassG <= 0.0) THEN
    _bParamBad := TRUE;                     // 目标量非法锁存 / Illegal target latched
END_IF
IF (fScaleMassG <> fScaleMassG) OR (ABS(fScaleMassG) > DL_DOS_INF) THEN
    _bScaleErr := TRUE;                     // 秤读数非有限归入秤异常（0319 复用，R90） / Non-finite scale folded into the scale fault
END_IF
IF (fCoarseFineKg < 0.0) OR (fCoarseFineKg > 1.0) THEN
    _bParamBad := TRUE;                     // 切换占比域外锁存 / Switch ratio out of range latched
END_IF
IF (tSettleTime <= T#0MS) OR (tSettleTime > DL_DOS_TO_WEIGH) THEN
    _bParamBad := TRUE;                     // 确认窗组态越界：为 0 或大于步 1 超时（结构性超时）锁存 / Confirm window out of range, latched
END_IF
IF xCoastAbort AND (tCoastTime <= T#0MS) THEN
    _bParamBad := TRUE;                     // 惰转窗组态越界：两段化中止永不收口锁存 / Coast window out of range, latched
END_IF

(*------------------------------------------------------------------------------
 * 段 4｜称重回退检测（注液执行期）：比上拍小超容差 → 0319 锁存
 *      Scale regression detection during the dosing execution phases
 *-----------------------------------------------------------------------------*)
IF (_ePhase = E_DL_ElyteDosingPhase.eCoarseFill)
   OR (_ePhase = E_DL_ElyteDosingPhase.eFineFill)
   OR (_ePhase = E_DL_ElyteDosingPhase.eSettle) THEN
    IF fScaleMassG < (_fScalePrevG - DL_DOS_TOL_G) THEN
        _bScaleErr := TRUE;                 // 称重回退锁存（暂停顺控保持输出） / Scale regression latched, sequencing paused
    END_IF
END_IF
_fScalePrevG := fScaleMassG;                // 快照推进 / Snapshot advanced

(*------------------------------------------------------------------------------
 * 段 5｜中止入口（任意拍生效；中止族态内不重复触发）与复位
 *      Abort entry, effective on any scan, not re-triggered in the family
 *-----------------------------------------------------------------------------*)
IF bAbort AND (_uAbortStage = 0)
   AND (_ePhase = E_DL_ElyteDosingPhase.eVacuumDraw
        OR _ePhase = E_DL_ElyteDosingPhase.eWeighCheck
        OR _ePhase = E_DL_ElyteDosingPhase.eCoarseFill
        OR _ePhase = E_DL_ElyteDosingPhase.eFineFill
        OR _ePhase = E_DL_ElyteDosingPhase.eSettle) THEN
    _uAbortStage := 1;                      // 进中止段 A（惰转） / Enter abort stage A, coast
END_IF
IF _uAbortStage >= 1 THEN
    IF (NOT bStart) AND (_uAbortStage = 2) THEN
        _uAbortStage := 0;                  // 关阀已完成且启动撤销，回空闲 / Close done and start dropped, back to idle
        _ePhase      := E_DL_ElyteDosingPhase.eIdle; // 相位回空闲 / Phase back to idle
    END_IF
END_IF
IF bReset THEN
    _bScaleErr := FALSE;                    // 复位清秤异常锁存 / Reset clears the scale latch
END_IF

(*------------------------------------------------------------------------------
 * 段 6｜四只计时无条件刷新（R40：CASE 之外每拍必调，各司其职不复用）
 *      Four timers refreshed unconditionally per R40
 *-----------------------------------------------------------------------------*)
fbDraw(IN := (_ePhase = E_DL_ElyteDosingPhase.eVacuumDraw) AND (_uAbortStage = 0),
       PT := DL_DOS_DRAW_T);               // 抽液计时 / Draw timer
fbStable(IN := (_ePhase = E_DL_ElyteDosingPhase.eWeighCheck) AND (_uAbortStage = 0)
              AND (ABS(fScaleMassG - _fBaseMassG) < DL_DOS_TOL_G), PT := tSettleTime); // 称重稳定窗 / Weigh stability window
fbSettle(IN := (_ePhase = E_DL_ElyteDosingPhase.eSettle) AND (_uAbortStage = 0), PT := tSettleTime); // 静置计时 / Settle timer
fbCoast(IN := (_uAbortStage = 1), PT := tCoastTime); // 中止惰转计时（段 A） / Abort coast timer, stage A

(*------------------------------------------------------------------------------
 * 段 7｜步进器单调用点（每拍恰好一次）与步完成判据装配
 *      Single sequencer call site and the step-done criteria assembly
 *-----------------------------------------------------------------------------*)
_bSeqStart := bStart AND (NOT _bStartPrev) AND (_ePhase = E_DL_ElyteDosingPhase.eIdle)
              AND (NOT _bParamBad) AND (NOT _bScaleErr); // 启动沿（空闲且组态合法） / Start edge in idle with a legal configuration
_bStartPrev := bStart;                      // 电平快照推进 / Level snapshot advanced

IF (_ePhase <> E_DL_ElyteDosingPhase.eIdle) AND (_ePhase <> E_DL_ElyteDosingPhase.eFault)
   AND (_uAbortStage = 0) THEN
    _abStepDone[0] := fbDraw.Q;             // 步 0 完成：抽液计时满 / Step 0 done, draw elapsed
    _abStepDone[1] := fbStable.Q;           // 步 1 完成：秤读数稳定窗满 / Step 1 done, stability window elapsed
    _abStepDone[2] := (fScaleMassG - _fBaseMassG) >= (fTargetMassG * fCoarseFineKg); // 步 2 完成：达粗细切换点 / Step 2 done, switch point reached
    _abStepDone[3] := (fScaleMassG - _fBaseMassG) >= fTargetMassG; // 步 3 完成：达目标量 / Step 3 done, target reached
    _abStepDone[4] := fbSettle.Q;           // 步 4 完成：静置计时满 / Step 4 done, settle elapsed
    _abStepDone[5] := TRUE;                 // 步 5 完成态恒成 / Step 5 always done
    IF _abStepDone[2] AND (_ePhase = E_DL_ElyteDosingPhase.eCoarseFill) THEN
        _bInfoCoarse := TRUE;               // 粗细切换点已达（信息级） / Switch point reached, info
    END_IF
END_IF

fbSeq(bStart := _bSeqStart, abStepDone := _abStepDone, auStepTimeout := _auStepTimeout,
      bHold := FALSE, bSingleStep := FALSE, bAdvance := FALSE,
      bAbort := (_uAbortStage >= 1), bReset := FALSE); // 步进器唯一调用点 / The only sequencer call site

IF _uAbortStage = 1 THEN
    IF fbCoast.Q THEN
        _uAbortStage := 2;                  // 惰转窗满，进中止段 B（关阀） / Coast elapsed, abort stage B, close
    END_IF
END_IF

(*------------------------------------------------------------------------------
 * 段 8｜相位机（只做迁移与步进对账；输出在段 9 按相置位）
 *      Phase machine, transitions and step reconciliation only
 *-----------------------------------------------------------------------------*)
CASE _ePhase OF

    E_DL_ElyteDosingPhase.eIdle:           // 空闲：启动沿锁定基线进抽液
        IF _bSeqStart THEN
            _fBaseMassG := fScaleMassG;     // 基线锁定 / Baseline locked
            _ePhase     := E_DL_ElyteDosingPhase.eVacuumDraw; // 进抽液相 / To the draw phase
        END_IF

    E_DL_ElyteDosingPhase.eVacuumDraw:     // 抽液：步进器推进到步 1 即转称重
        IF fbSeq.bError THEN
            _ePhase := E_DL_ElyteDosingPhase.eFault; // 步超时，故障 / Step timeout, fault
        ELSIF (fbSeq.nCurrentStep = 1) THEN
            _ePhase := E_DL_ElyteDosingPhase.eWeighCheck; // 步进器已推进 / The sequencer advanced
        END_IF

    E_DL_ElyteDosingPhase.eWeighCheck:     // 称重核对：步进器推进到步 2 即转粗注
        IF fbSeq.bError THEN
            _ePhase := E_DL_ElyteDosingPhase.eFault; // 步超时，故障 / Step timeout, fault
        ELSIF (fbSeq.nCurrentStep = 2) THEN
            _ePhase := E_DL_ElyteDosingPhase.eCoarseFill; // 步进器已推进 / The sequencer advanced
        END_IF

    E_DL_ElyteDosingPhase.eCoarseFill:     // 粗注：步进器推进到步 3 即转细注
        IF fbSeq.bError THEN
            _ePhase := E_DL_ElyteDosingPhase.eFault; // 步超时，故障 / Step timeout, fault
        ELSIF (fbSeq.nCurrentStep = 3) THEN
            _ePhase := E_DL_ElyteDosingPhase.eFineFill; // 步进器已推进 / The sequencer advanced
        END_IF

    E_DL_ElyteDosingPhase.eFineFill:       // 细注：步进器推进到步 4 即转静置
        IF fbSeq.bError THEN
            _ePhase := E_DL_ElyteDosingPhase.eFault; // 步超时，故障 / Step timeout, fault
        ELSIF (fbSeq.nCurrentStep = 4) THEN
            _ePhase := E_DL_ElyteDosingPhase.eSettle; // 步进器已推进 / The sequencer advanced
        END_IF

    E_DL_ElyteDosingPhase.eSettle:         // 静置：步进器推进到步 5 即完成
        IF fbSeq.bError THEN
            _ePhase := E_DL_ElyteDosingPhase.eFault; // 步超时，故障 / Step timeout, fault
        ELSIF (fbSeq.nCurrentStep = 5) THEN
            _ePhase := E_DL_ElyteDosingPhase.eDone; // 步进器已推进 / The sequencer advanced
        END_IF

    E_DL_ElyteDosingPhase.eDone:           // 完成：等启动撤销回空闲
        IF NOT bStart THEN
            _ePhase := E_DL_ElyteDosingPhase.eIdle; // 回空闲 / Back to idle
        END_IF

    E_DL_ElyteDosingPhase.eFault:          // 故障：复位沿且原因消失回空闲
        IF bReset AND (NOT _bParamBad) AND (NOT _bScaleErr) THEN
            _ePhase := E_DL_ElyteDosingPhase.eIdle; // 回空闲 / Back to idle
        END_IF

    ELSE                                   // 非法状态兜底（R21：CASE 必带 ELSE）
        _bIllegal := TRUE;                 // 标记非法状态 / Flag the illegal state
        _ePhase   := E_DL_ElyteDosingPhase.eFault; // 回故障态（段 9 全断） / Back to fault, all outputs off
END_CASE

(*------------------------------------------------------------------------------
 * 段 9｜输出置位（次序即安全：泵先于阀；中止段 A 泵断使能、阀保持不动，
 *       机检断言：abort 拍不得出现关阀输出置位——段 A 阀输出 = 保持量）
 *      Output assignment, pump precedes the valve, abort stage A holds the valve
 *-----------------------------------------------------------------------------*)
CASE _ePhase OF
    E_DL_ElyteDosingPhase.eVacuumDraw:     // 抽液：泵运行 / Draw: pump runs
        bPumpOut := (_uAbortStage = 0);    // 中止段 A 泵使能立即断 / Pump enable cut immediately in abort stage A
    E_DL_ElyteDosingPhase.eCoarseFill:     // 粗注：阀开 / Coarse: valve open
        bDosingOut := (_uAbortStage = 0) OR (_uAbortStage = 1); // 段 A 阀保持，段 B 关阀 / Valve held in stage A, closed in stage B
    E_DL_ElyteDosingPhase.eFineFill:       // 细注：阀开 / Fine: valve open
        bDosingOut := (_uAbortStage = 0) OR (_uAbortStage = 1); // 段 A 阀保持，段 B 关阀 / Valve held in stage A, closed in stage B
    ELSE                                   // 其余相输出全断 / Otherwise all off
        bDosingOut := FALSE;               // 注液阀断 / Dosing off
        bPumpOut   := FALSE;               // 泵断 / Pump off
END_CASE
IF (NOT xCoastAbort) AND (_uAbortStage >= 1) THEN
    bDosingOut := FALSE;                   // 兼容路径：单拍中止（不推荐，残压回流风险） / Legacy single-scan abort, not recommended
    bPumpOut   := FALSE;                   // 泵同拍断 / Pump off the same scan
END_IF

fDosedMassG := fScaleMassG - _fBaseMassG;   // 已注量出口 [克] / Dosed mass outlet [g]
IF fDosedMassG < 0.0 THEN
    fDosedMassG := 0.0;                     // 负增量钳 0（换批/去皮期） / Negative delta clamped to zero
END_IF
ePhase := _ePhase;                          // 相位出口 / Phase outlet

IF _bIllegal THEN
    eErr   := 16#0005_031A;                 // 故障级：状态机兜底 / Fault: state machine fallback
    bError := TRUE;                         // 置故障标志 / Raise the fault flag
ELSIF _bParamBad THEN
    eErr   := 16#0005_0318;                 // 故障级：目标量或占比非法 / Fault: illegal target or ratio
    bError := TRUE;                         // 置故障标志 / Raise the fault flag
ELSIF _bScaleErr THEN
    eErr   := 16#0005_0319;                 // 故障级：称重回退判秤异常 / Fault: scale regression
    bError := TRUE;                         // 置故障标志 / Raise the fault flag
ELSIF fbSeq.bError THEN
    eErr   := 16#0005_031A;                 // 故障级：步超时复用兜底码（R90） / Fault: step timeout, code reused per R90
    bError := TRUE;                         // 置故障标志 / Raise the fault flag
ELSIF _bInfoCoarse THEN
    eErr := 16#0005_01E2;                   // 信息级：粗细切换点已达 / Info: switch point reached
END_IF

bValid := (NOT bError) AND (_ePhase <> E_DL_ElyteDosingPhase.eIdle); // 空闲/故障输出不可用 / Outputs unusable in idle or fault
END_FUNCTION_BLOCK

(* ---- FB_DL_ElectrolyteDosingTrend.st ---- *)
(*
  ==================================================================
  组件名 Component  : FB_DL_ElectrolyteDosingTrend
  分类   Category   : DL_Process
  版本   Version    : 1.0.0
  功能   Purpose    : 注液量趋势 SPG（统计过程判据）统计。逐次注液量进环窗，
                      窗满后给出均值、样本标准差、上下控制限（均值 ± k × 标准差）、
                      越限判据与连续同向趋势判据（连升 / 连降），并给目标带内
                      合格判据，用于注液泵磨损与堵塞的早期趋势预警。
  溯源   Origin     : 均值 / 标准差 / 控制限为公开统计过程控制口径；本件为 clean-room
                      实现，仅借鉴来源分类与参数域组织（来源标签 roadmap-p2-dosing），
                      道莅原创设计，未复制任何闭源代码行。
  平台   Platform   : 纯 IEC 61131-3（SQRT / REAL / R_TRIG，无私有库、无方言转换）
  作者   Author     : 道莅代码库 · PLC 编程专家（R55）
  ------------------------------------------------------------------
  边界 Boundary     :
                      一 本件只做统计与趋势判据，不调节注液泵、不改配方（属主边界）；
                      二 样本标准差按 n − 1 无偏口径，样本数小于 2 时不下结论；
                      三 方差由「平方和 − 和的平方 / n」推得，舍入致负值一律钳零（开方前闸）；
                      四 环窗遍历按时间序遍历，禁按数组下标序遍历（R194）；
                      五 无全局变量、无外部变量声明、无物理地址寻址。
  输出契约 Output contract:
                      fMeanMl / fStdMl / fUclMl / fLclMl 仅在样本数达标时更新，
                      否则保持上拍值；bOutOfCtrl 仅在最新样本越限时为真（单拍语义，
                      由调用方按需累计）；nTrendRun 正数为连升、负数为连降；
                      eCause 故障级成因与 bError 配对（R45），信息级永不置 bError。
  修订记录 Revision  :
    2026-11-20  v1.0.0  R55 首版（批 4 · 序号 15）
  ==================================================================
*)

TYPE E_DL_EdtTrend :
(
    eStable := 0,       // 平稳：最新与上一样本无明显方向 / stable, no clear direction between the last two samples
    eUp     := 10,      // 连升：连续同向上升 / rising, a run of increases
    eDown   := 20       // 连降：连续同向下降 / falling, a run of decreases
);
END_TYPE

TYPE E_DL_EdtCause :
(
    eNone       := 0,   // 无成因 / no cause
    eCfgIllegal := 1,   // 组态非法：窗口容量、系数或目标带越域（故障级，与 bError 配对）/ illegal config, window size, sigma factor or target band out of domain
    eNoSample   := 2,   // 样本数不足 2，统计量保持上拍值（信息级）/ fewer than two samples and the statistics hold, informational
    eBadSample  := 3    // 存在非有限样本，已拒收（信息级）/ non-finite samples were rejected, informational
);
END_TYPE

FUNCTION_BLOCK FB_DL_ElectrolyteDosingTrend
VAR_INPUT
    bEnable      : BOOL := TRUE;             // 使能，失能时不收样本 [-] / enable, no sample is accepted when disabled
    bReset       : BOOL := FALSE;           // 复位上升沿清故障锁存与全部统计 [-] / reset rising edge clears the fault latch and all statistics
    bSamplePulse : BOOL := FALSE;            // 单次注液量采样脉冲，上升沿收一条 [-] / single dose sample pulse, one sample per rising edge
    fVolMl       : REAL := 0.0;              // 本次注液量 [毫升] / dose volume of this shot [millilitre]
    fTargetMl    : REAL := 100.0;            // 目标注液量 [毫升]，域 大于零 / target dose volume [millilitre], domain above zero
    fTolPct      : REAL := 2.0;              // 目标带容差 [百分比]，域 大于零 / target band tolerance [percent], domain above zero
    nWinSize     : INT := 20;                // 统计窗样本数 [个]，域 2..64 / statistics window size [count], domain 2 to 64
    fSigmaK      : REAL := 3.0;              // 控制限系数（倍标准差）[倍]，域 1..6 / control limit factor in standard deviations [factor], domain 1 to 6
END_VAR
VAR_OUTPUT
    fMeanMl      : REAL := 0.0;              // 窗口均值 [毫升] / window mean [millilitre]
    fStdMl       : REAL := 0.0;              // 窗口样本标准差（n − 1 口径）[毫升] / window sample standard deviation over n minus one [millilitre]
    fUclMl       : REAL := 0.0;              // 上控制限 [毫升] / upper control limit [millilitre]
    fLclMl       : REAL := 0.0;              // 下控制限 [毫升]，可为负 / lower control limit, may be negative [millilitre]
    nSampleCnt   : INT := 0;                 // 窗口有效样本数 [个] / valid sample count in the window
    bOutOfCtrl   : BOOL := FALSE;            // 最新样本越控制限 [-] / the newest sample is beyond a control limit
    bHasStats    : BOOL := FALSE;            // 统计量是否已可交付 [-] / the statistics are deliverable
    bInTarget    : BOOL := FALSE;            // 最新样本落在目标带内 [-] / the newest sample is inside the target band
    nTrendRun    : INT := 0;                 // 连续同向计数（正连升 / 负连降）[次] / signed run length, positive rising and negative falling [count]
    eTrend       : E_DL_EdtTrend := E_DL_EdtTrend.eStable; // 趋势出口 [枚举] / trend outlet [enum]
    nRejectCnt   : INT := 0;                 // 累计拒收样本数（饱和到上限）[个] / total rejected samples, saturated [count]
    eCause       : E_DL_EdtCause := E_DL_EdtCause.eNone; // 成因出口 [枚举] / cause outlet [enum]
    bError       : BOOL := FALSE;            // 故障锁存标志 [-] / fault latch flag
END_VAR
VAR
    rtSample     : R_TRIG;                   // 采样沿检测，段 0 无条件刷新 / sample edge detector, refreshed unconditionally in segment zero
    rtReset      : R_TRIG;                   // 复位沿检测，段 0 无条件刷新 / reset edge detector, refreshed unconditionally in segment zero
    _eCause      : E_DL_EdtCause := E_DL_EdtCause.eNone;  // 信息级成因，每拍重算 / informational cause, recomputed every scan
    _eFaultCause : E_DL_EdtCause := E_DL_EdtCause.eNone;  // 故障级成因，锁存至复位沿 / fault cause, latched until the reset edge
    _eTrend      : E_DL_EdtTrend := E_DL_EdtTrend.eStable; // 趋势工作值 / trend working value
    _bFault      : BOOL := FALSE;            // 故障锁存位 [-] / fault latch bit
    _bInit       : BOOL := FALSE;            // 首扫初始化完成标志（R310）/ first scan initialisation flag
    _bCfgBad     : BOOL := FALSE;            // 组态非法判定 [-] / illegal configuration verdict
    _bSampleOk   : BOOL := FALSE;            // 本拍样本有限 [-] / this scan sample finite
    _bStatsOk    : BOOL := FALSE;            // 统计量可算 [-] / the statistics are computable
    _bVarOk      : BOOL := FALSE;            // 方差非负可开方 [-] / the variance is non-negative and can be rooted
    _bBadReject  : BOOL := FALSE;            // 本拍发生过拒收 [-] / a rejection occurred this scan
    _nWinUse     : INT := 2;                 // 钳定后的窗口容量 [个] / clamped window size [count]
    _nFill       : INT := 0;                 // 环窗已填样本数 [个] / samples held in the ring [count]
    _nHead       : INT := 0;                 // 环窗最新样本槽位（1 起，回钳 1..64）[槽号] / newest ring slot, clamped one through sixty four
    _nIdx        : INT := 0;                 // 环窗游标 [槽号] / ring cursor [slot]
    _nK          : INT := 0;                 // 时间序遍历序号 [序号] / time-order ordinal
    _nGuard      : INT := 0;                 // 遍历守护计数 [次] / traversal guard [count]
    _nRun        : INT := 0;                 // 连续同向计数工作值 [次] / signed run length working value [count]
    _nReject     : INT := 0;                 // 拒收计数工作值 [个] / rejected sample count [count]
    _fVolPrev    : REAL := 0.0;              // 上一样本注液量 [毫升] / previous sample volume [millilitre]
    _fSum        : REAL := 0.0;              // 窗口和 [毫升] / window sum [millilitre]
    _fSumSq      : REAL := 0.0;              // 窗口平方和 [毫升平方] / window sum of squares [millilitre squared]
    _fMean       : REAL := 0.0;              // 均值工作值 [毫升] / mean working value [millilitre]
    _fVar        : REAL := 0.0;              // 方差工作值 [毫升平方] / variance working value [millilitre squared]
    _fStd        : REAL := 0.0;              // 标准差工作值 [毫升] / standard deviation working value [millilitre]
    _fDivN       : REAL := 1.0;              // 均值除子（样本数）[个] / mean divisor, the sample count [count]
    _fDivNm1     : REAL := 1.0;              // 方差除子（样本数减一）[个] / variance divisor, the sample count minus one [count]
    _fVolLoc     : REAL := 0.0;              // 遍历取出的样本值 [毫升] / sample value taken during the traversal [millilitre]
    _afVol       : ARRAY[1..64] OF REAL := [64(0.0)]; // 环窗注液量缓存 [毫升] / ring buffer of dose volumes [millilitre]
END_VAR
VAR CONSTANT
    DL_EDT_MAX       : INT := 64;            // 环窗容量与槽位回钳上界 [个] / ring capacity and slot clamp upper bound
    DL_EDT_WIN_MIN   : INT := 2;             // 窗口容量下限（标准差至少两个样本）[个] / window size floor, a deviation needs two samples
    DL_EDT_VOL_MAX   : REAL := 1.0E6;        // 注液量量级上限，防量纲错配 [毫升] / dose volume magnitude ceiling against a mismatch [millilitre]
    DL_EDT_SIGMA_MIN : REAL := 1.0;          // 控制限系数下限 [倍] / control limit factor floor [factor]
    DL_EDT_SIGMA_MAX : REAL := 6.0;          // 控制限系数上限 [倍] / control limit factor ceiling [factor]
    DL_EDT_TOL_MAX   : REAL := 100.0;        // 容差上限 [百分比] / tolerance ceiling [percent]
    DL_EDT_REJ_MAX   : INT := 30000;         // 拒收计数上限，防溢出 [个] / rejection count ceiling against overflow [count]
    DL_EDT_VAR_EPS   : REAL := 1.0E-9;       // 方差零阈，舍入负值钳零用 [毫升平方] / variance zero threshold for clamping rounding negatives [millilitre squared]
END_VAR

// 段 0｜沿检测无条件周期刷新（禁入分支）/ segment 0, unconditional refresh of the edge detectors, never inside a branch
rtSample(CLK := bSamplePulse); // 采样沿无条件刷新 / unconditional refresh of the sample edge
rtReset(CLK := bReset); // 复位沿无条件刷新 / unconditional refresh of the reset edge

// 段 1｜首扫初始化（R310）/ segment 1, first scan initialisation
IF NOT _bInit THEN // 首扫一拍 / the very first scan
    _bInit := TRUE; // 置首扫完成标志 / raise the first scan flag
    _bFault := FALSE; // 故障锁存清零 / clear the fault latch
    _eCause := E_DL_EdtCause.eNone; // 信息级成因清零 / clear the informational cause
    _eFaultCause := E_DL_EdtCause.eNone; // 故障级成因清零 / clear the fault cause
    _nHead := 0; // 环窗无样本 / the ring holds no sample
    _nFill := 0; // 环窗计数清零 / clear the ring count
    _nRun := 0; // 趋势计数清零 / clear the run counter
    _fVolPrev := 0.0; // 上一样本清零 / clear the previous sample
    _eTrend := E_DL_EdtTrend.eStable; // 趋势从平稳起步 / the trend starts stable
END_IF

// 段 2｜复位沿作用域：清锁存 / 清统计 / 清环窗游标（三项逐项声明）/ segment 2, reset edge scope
IF rtReset.Q THEN // 复位沿 / reset edge
    _bFault := FALSE; // 作用域一：清故障锁存 / scope one, clear the fault latch
    _eFaultCause := E_DL_EdtCause.eNone; // 作用域一：清故障级成因 / scope one, clear the fault cause
    _nHead := 0; // 作用域三：清环窗槽位 / scope three, clear the ring slot cursor
    _nFill := 0; // 作用域三：清环窗计数 / scope three, clear the ring count
    _nRun := 0; // 作用域二：清趋势计数 / scope two, clear the run counter
    _nReject := 0; // 作用域二：清拒收计数 / scope two, clear the rejection count
    _fVolPrev := 0.0; // 作用域二：清上一样本 / scope two, clear the previous sample
    _eTrend := E_DL_EdtTrend.eStable; // 作用域二：趋势回平稳 / scope two, the trend returns to stable
    fMeanMl := 0.0; // 作用域二：清均值出口 / scope two, clear the mean outlet
    fStdMl := 0.0; // 作用域二：清标准差出口 / scope two, clear the deviation outlet
    fUclMl := 0.0; // 作用域二：清上控制限出口 / scope two, clear the upper limit outlet
    fLclMl := 0.0; // 作用域二：清下控制限出口 / scope two, clear the lower limit outlet
END_IF

// 段 3｜组态域闸（R151 全覆盖）/ segment 3, configuration domain gate over every pin
_bCfgBad := FALSE; // 组态非法预置假 / preset the illegal configuration verdict to false
IF (fTargetMl <= 0.0) OR (fTargetMl <> fTargetMl) OR (fTargetMl > DL_EDT_VOL_MAX) THEN // 目标量越域 / the target is out of domain
    _bCfgBad := TRUE; // 判非法 / mark illegal
END_IF
IF (fTolPct <= 0.0) OR (fTolPct > DL_EDT_TOL_MAX) OR (fTolPct <> fTolPct) THEN // 容差越域 / the tolerance is out of domain
    _bCfgBad := TRUE; // 判非法 / mark illegal
END_IF
IF (nWinSize < DL_EDT_WIN_MIN) OR (nWinSize > DL_EDT_MAX) THEN // 窗口容量越域 / the window size is out of domain
    _bCfgBad := TRUE; // 判非法 / mark illegal
END_IF
IF (fSigmaK < DL_EDT_SIGMA_MIN) OR (fSigmaK > DL_EDT_SIGMA_MAX) OR (fSigmaK <> fSigmaK) THEN // 系数越域 / the factor is out of domain
    _bCfgBad := TRUE; // 判非法 / mark illegal
END_IF
IF _bCfgBad AND (NOT _bFault) THEN // 组态非法且未锁存 / illegal configuration and not yet latched
    _bFault := TRUE; // 置故障锁存 / raise the fault latch
    _eFaultCause := E_DL_EdtCause.eCfgIllegal; // 故障级成因 (R45 配对 bError) / fault grade cause paired with bError
END_IF
_nWinUse := nWinSize; // 窗口容量直通 / the window size passes through
IF _nWinUse < DL_EDT_WIN_MIN THEN // 下越界 / below the lower bound
    _nWinUse := DL_EDT_WIN_MIN; // 回钳到 2 / clamp to two
ELSIF _nWinUse > DL_EDT_MAX THEN // 上越界 / above the upper bound
    _nWinUse := DL_EDT_MAX; // 回钳到 64 / clamp to sixty four
END_IF

// 段 4｜样本接收与趋势跟踪 / segment 4, sample acceptance and trend tracking
_eCause := E_DL_EdtCause.eNone; // 信息级成因每拍重算 / the informational cause is recomputed every scan
_bBadReject := FALSE; // 拒收标志预置假 / preset the rejection flag to false
IF rtSample.Q AND bEnable AND (NOT _bFault) THEN // 采样沿且使能无故障 / sample edge while enabled and unfaulted
    _bSampleOk := (fVolMl = fVolMl) AND ((fVolMl - fVolMl) = (fVolMl - fVolMl)) AND (fVolMl >= 0.0) AND (fVolMl <= DL_EDT_VOL_MAX); // 样本有限性与量级闸 / sample finiteness and magnitude gate
    IF NOT _bSampleOk THEN // 样本不可用 / the sample is unusable
        _bBadReject := TRUE; // 记拒收 / record the rejection
        IF _nReject < DL_EDT_REJ_MAX THEN // 未达计数上限 / below the ceiling
            _nReject := _nReject + 1; // 拒收计数递增 / increment the rejection count
        END_IF
    ELSE
        // 段 4.1｜环窗写入：先算槽位再写入，槽位回钳 1..64 / segment 4.1, ring write with a clamped slot
        _nHead := _nHead + 1; // 槽位前移 / advance the slot
        IF _nHead > DL_EDT_MAX THEN // 越过上界 / past the upper bound
            _nHead := 1; // 回钳到一号槽 / clamp back to slot one
        END_IF
        _afVol[_nHead] := fVolMl; // 样本入环窗 / store the sample
        IF _nFill < DL_EDT_MAX THEN // 环窗未满 / the ring is not yet full
            _nFill := _nFill + 1; // 计数递增 / increment the count
        END_IF
        // 段 4.2｜趋势跟踪：与上一样本比较方向 / segment 4.2, trend tracking against the previous sample
        IF _nFill > 1 THEN // 至少两条样本才有方向 / a direction needs at least two samples
            IF fVolMl > _fVolPrev THEN // 上升 / rising
                IF _nRun < 0 THEN // 原为连降 / previously falling
                    _nRun := 1; // 方向翻转，计数从 1 起 / the direction flipped and the run restarts at one
                ELSE
                    _nRun := _nRun + 1; // 连升累加 / extended the rising run
                END_IF
            ELSIF fVolMl < _fVolPrev THEN // 下降 / falling
                IF _nRun > 0 THEN // 原为连升 / previously rising
                    _nRun := -1; // 方向翻转，计数从负 1 起 / the direction flipped and the run restarts at minus one
                ELSE
                    _nRun := _nRun - 1; // 连降累加 / extended the falling run
                END_IF
            ELSE // 相等（本拍样本与上一样本同值）/ equal to the previous sample
                _nRun := 0; // 无方向 / no direction
            END_IF
        END_IF
        _fVolPrev := fVolMl; // 上一样本推进 / advance the previous sample
    END_IF
END_IF
IF _bBadReject THEN // 本拍发生拒收 / a rejection occurred this scan
    _eCause := E_DL_EdtCause.eBadSample; // 信息级成因 / informational cause
END_IF

// 段 5｜统计量：按时间序遍历环窗求均值与样本标准差 / segment 5, statistics over the ring in time order
_bStatsOk := _nFill >= DL_EDT_WIN_MIN; // 样本数达下限才可算标准差 / the deviation needs the minimum sample count
IF _bStatsOk THEN // 统计可算 / the statistics are computable
    _fSum := 0.0; // 和清零 / clear the sum
    _fSumSq := 0.0; // 平方和清零 / clear the sum of squares
    _nIdx := _nHead - _nFill + 1; // 时间序最旧槽位 / the oldest slot in time order
    IF _nIdx < 1 THEN // 越过下界 / below the lower bound
        _nIdx := _nIdx + DL_EDT_MAX; // 单次回绕补齐 / a single wrap restores the time order
    END_IF
    _nK := 1; // 时间序序号自 1 起 / the time-order ordinal starts at one
    _nGuard := 0; // 守护计数清零 / reset the guard
    WHILE (_nK <= _nFill) AND (_nGuard < (2 * DL_EDT_MAX)) DO // 双重守护 / dual guard
        _nGuard := _nGuard + 1; // 守护计数递增 / increment the guard
        _nIdx := _nHead - _nFill + _nK; // 时间序槽位 / the slot in time order
        IF _nIdx < 1 THEN // 越过下界 / below the lower bound
            _nIdx := _nIdx + DL_EDT_MAX; // 单次回绕 / single wrap
        END_IF
        _fVolLoc := _afVol[_nIdx]; // 取出样本 / take the sample
        _fSum := _fSum + _fVolLoc; // 累加和 / accumulate the sum
        _fSumSq := _fSumSq + _fVolLoc * _fVolLoc; // 累加平方和 / accumulate the sum of squares
        _nK := _nK + 1; // 序号递增 / increment the ordinal
    END_WHILE
    _fDivN := INT_TO_REAL(_nFill); // 均值除子为样本数，已证不小于 2 / the mean divisor is the count, proven not below two
    _fMean := _fSum / _fDivN; // 均值 / mean
    _fDivNm1 := INT_TO_REAL(_nFill - 1); // 方差除子为 n − 1，已证不小于 1 / the variance divisor is n minus one, proven not below one
    _fVar := (_fSumSq - (_fSum * _fSum) / _fDivN) / _fDivNm1; // 无偏方差 / unbiased variance
    _bVarOk := _fVar > DL_EDT_VAR_EPS; // 方差可用（舍入负值不参与开方）/ the variance is usable and rounding negatives are excluded
    IF _bVarOk THEN // 方差可用 / the variance is usable
        _fStd := SQRT(_fVar); // 标准差 / standard deviation
    ELSE
        _fStd := 0.0; // 方差近零时标准差记零 / a near-zero variance yields a zero deviation
    END_IF
    fMeanMl := _fMean; // 均值出口 / mean outlet
    fStdMl := _fStd; // 标准差出口 / deviation outlet
    fUclMl := _fMean + fSigmaK * _fStd; // 上控制限 / upper control limit
    fLclMl := _fMean - fSigmaK * _fStd; // 下控制限（可为负）/ lower control limit, may be negative
    bHasStats := TRUE; // 统计量可交付 / the statistics are deliverable
ELSE // 样本不足 / too few samples
    bHasStats := FALSE; // 统计量不可交付，出口保持上拍值 / the statistics are not deliverable and the outlets hold
    _eCause := E_DL_EdtCause.eNoSample; // 信息级成因 / informational cause
END_IF

// 段 6｜越限与目标带判据（仅在有统计量时判，避免用未成型的限值下结论）/ segment 6, limit and target band verdicts
bOutOfCtrl := FALSE; // 越限标志预置假 / preset the out-of-control flag to false
bInTarget := FALSE; // 目标带标志预置假 / preset the in-target flag to false
IF bHasStats AND rtSample.Q AND _bSampleOk THEN // 仅在有效采样拍判越限与目标带 / the verdicts run only on a valid sample scan
    bOutOfCtrl := (fVolMl > fUclMl) OR (fVolMl < fLclMl); // 最新样本越控制限 / the newest sample is beyond a control limit
    bInTarget := ABS(fVolMl - fTargetMl) <= (fTargetMl * fTolPct / 100.0); // 目标带判据，除子为常量 100.0 / target band verdict with the constant divisor one hundred
END_IF

// 段 7｜趋势出口映射 / segment 7, trend outlet mapping
IF _nRun > 0 THEN // 连升 / rising run
    _eTrend := E_DL_EdtTrend.eUp; // 连升档 / rising
ELSIF _nRun < 0 THEN // 连降 / falling run
    _eTrend := E_DL_EdtTrend.eDown; // 连降档 / falling
ELSE
    _eTrend := E_DL_EdtTrend.eStable; // 平稳档 / stable
END_IF
eTrend := _eTrend; // 趋势出口单点映射 / single-point trend outlet mapping
nTrendRun := _nRun; // 连续同向计数出口 / signed run length outlet
nSampleCnt := _nFill; // 窗口样本数出口 / window sample count outlet
nRejectCnt := _nReject; // 拒收计数出口 / rejection count outlet
IF _bFault THEN // 故障锁存优先 / the fault latch takes priority
    eCause := _eFaultCause; // 故障级成因锁存回放 / the fault cause is replayed from the latch
ELSE
    eCause := _eCause; // 信息级成因直映 / the informational cause is mapped directly
END_IF
bError := _bFault; // 故障标志与锁存位同源 / the fault flag shares the latch source
END_FUNCTION_BLOCK

(* ---- FB_DL_ElectrolyteFillCtrl.st ---- *)
(*
  FB_DL_ElectrolyteFillCtrl  —  注液量闭环（称重罐减量法 + 静置浸润计时）/ Electrolyte fill closed loop, mass-loss method
  分类 Category : DL_Process
  码位 Code     : 16#06_0_B7
  段位说明      : B6 格由 HjtPvdSeq 启用，本件启用相邻 B7 格（一件一码）
  版本 Version  : 1.0.0
  来源 Source   : t2-2-lbp — 注液闭环工艺待挖项
  溯源 Origin   : clean-room 实现，减量法注液公开工艺语义借鉴，未复制任何源码行
                  （与 FB_DL_ElectrolyteDosingSeq 分工：那件是定量投加顺控，本件是减量法闭环注液 + 浸润驻留）
  功能 Function : 1) 六相顺控 Idle→Tare→Fill→Trim→Dwell→Done：皮重稳定采集 → 大流量粗注 →
                  微调收口 → 静置浸润驻留 → 完成；
                  2) 减量法口径：注液量 fFilledKg = 皮重 − 实时称重（罐在秤上，质量递减）；
                  3) 粗注→微调切换：剩余量经 FC_DL_Hysteresis 迟滞判入预关带（防阀门口径切换抖动）；
                  4) 收口判定：FB_DL_ToleranceWindow 三态判定注液量入容差 → 关阀进静置；
                  5) 静置浸润：tDwellTime 驻留，质量漂移超 fDwellDriftKg 置信息级码（渗漏提示不置故障）。
  边界 Boundary : ① 称重信号 fTankMassKg 非有限保持上次有效值；注液期质量上升（反流）判故障级锁存；
                  ② 组态域闸覆盖全部参与换算引脚（R151）；容差/提前量/驻留时长域非法判组态错；
                  ③ R228-A 达标声明：tonTareTo/tonFillTo/tonTrimTo/tonDwell 各自单相独占
                  （IN 为单相等式），跨相迁移拍 IN 必断；tonDwell PT 接浸润时长（配方语义）；
                  ④ R228-B 达标声明：eFault 迁出 = rtReset.Q（输入引脚，恒可达），逐字写于此；
                  ⑤ 阀门指令为开度百分比（rValveCmdPct），不写物理 IO（由上层 PRG_IoMapping 承载）；
                  ⑥ CASE 全态覆盖 + ELSE 兜底置 Fault。
  依赖 Depends  : FB_DL_ToleranceWindow / FB_DL_SignalStatistics（实例化，引脚按 registry 实名）；
                  FC_DL_Hysteresis（函数调用，bState 由本件成员持有回传）
  码表 Error codes（本件格 06_0_B7，子码步进 +0x100）:
    16#0006_01B7 信息级：注液周期完成（Done 相）
    16#0006_02B7 故障级：组态非法（目标/容差/提前量/漂移阈/驻留/超时域非法），锁存至复位
    16#0006_03B7 故障级：相超时（Tare/Fill/Trim 独立计时），锁存至复位
    16#0006_04B7 故障级：称重信号非有限持续 / 注液期质量上升（反流），锁存至复位
    16#0006_05B7 故障级：状态机落 ELSE 兜底（非法相位 ID）
    16#0006_06B7 信息级：静置期质量漂移超阈（渗漏提示，不置故障）
    16#0006_07B7 信息级：皮重稳定判据等待中（Tare 相，不置故障）

  修订历史 Revision :
    2026-11-19  v1.0.0  R39 首版（批次 3 · 序号 15）
*)

TYPE E_DL_ElytFillState :
(
    eIdle  := 0,    // 空闲：等启动指令 / Idle, waiting for start
    eTare  := 10,   // 皮重相：称重稳定后锁皮重 / Tare, lock tare after mass stable
    eFill  := 20,   // 粗注相：阀全开大流量 / Bulk fill, valve wide open
    eTrim  := 30,   // 微调相：收口至容差带 / Trim, close into tolerance band
    eDwell := 40,   // 静置相：浸润驻留 + 漂移监视 / Dwell, soaking with drift watch
    eDone  := 50,   // 完成：周期落定 / Done
    eFault := 90    // 故障：组态/超时/称重锁定 / Fault, latched
);
END_TYPE

FUNCTION_BLOCK FB_DL_ElectrolyteFillCtrl
VAR_INPUT
    bStart        : BOOL := FALSE;      // 启动指令（上升沿）/ Start command
    fTankMassKg   : REAL := 0.0;        // 称重罐实时质量 [kg] / Live tank mass from scale
    fBatchTargetKg: REAL := 5.0;        // 目标注液量 [kg]，域 > 0 / Target fill mass
    fFillTolKg    : REAL := 0.02;       // 注液量容差半宽 [kg]，域 > 0 / Fill tolerance half band
    fPrefillKg    : REAL := 0.10;       // 粗注→微调预关提前量 [kg]，域 > 0 / Pre-close lead mass
    fHystKg       : REAL := 0.02;       // 切换迟滞带 [kg]，域 > 0 / Switch hysteresis band
    fStatTolKg    : REAL := 0.005;      // 皮重/静置稳定峰峰阈 [kg]，域 > 0 / Stability peak-to-peak threshold
    fDwellDriftKg : REAL := 0.01;       // 静置漂移报警阈 [kg]，域 > 0 / Dwell drift alarm threshold
    tTareTo       : TIME := T#10S;      // 皮重相超时 [ms]，域 > 0 / Tare timeout
    tFillTo       : TIME := T#120S;     // 粗注相超时 [ms]，域 > 0 / Bulk fill timeout
    tTrimTo       : TIME := T#60S;      // 微调相超时 [ms]，域 > 0 / Trim timeout
    tDwellTime    : TIME := T#30S;      // 静置浸润时长 [ms]，域 > 0 / Dwell soaking duration
    bReset        : BOOL := FALSE;      // 复位（eFault 迁出唯一沿）/ Reset, sole fault exit edge
END_VAR
VAR_OUTPUT
    rValveCmdPct  : REAL;               // 注液阀开度指令 [%]（上层消费）/ Fill valve command output
    fFilledKg     : REAL;               // 已注液量 [kg] = 皮重 − 实时质量 / Filled mass by mass loss
    fRemainingKg  : REAL;               // 剩余注液量 [kg] / Remaining fill mass
    fTareKg       : REAL;               // 锁定皮重 [kg] / Locked tare mass
    bFillDone     : BOOL;               // 注液完成 / Fill cycle done
    bDwellDone    : BOOL;               // 静置浸润完成 / Dwell done
    nErrId        : UDINT;              // 事件码，0 = 无事件 / Event code
    eState        : E_DL_ElytFillState; // 状态出口，段尾单点映射 / State outlet
END_VAR
VAR
    fbTol      : FB_DL_ToleranceWindow; // 容差窗判定实例（主体首部无条件刷新）/ Tolerance window instance
    fbStat     : FB_DL_SignalStatistics;// 质量稳定统计窗实例（主体首部无条件刷新）/ Mass statistics window instance
    tonTareTo  : TON;                  // 皮重相超时（单相独占）/ Tare timeout, single phase
    tonFillTo  : TON;                  // 粗注相超时（单相独占）/ Bulk fill timeout, single phase
    tonTrimTo  : TON;                  // 微调相超时（单相独占）/ Trim timeout, single phase
    tonDwell   : TON;                  // 静置浸润计时（单相独占，PT=浸润时长）/ Dwell timer, single phase
    rtStart    : R_TRIG;               // 启动上升沿 / Start rising edge
    rtReset    : R_TRIG;               // 复位上升沿 / Reset rising edge
    _eState    : E_DL_ElytFillState := E_DL_ElytFillState.eIdle;   // 内部相位（CASE 唯一写入目标）/ Internal phase
    _rMassEff  : REAL;                 // 生效质量 [kg]（非有限保持载体）/ Effective mass with hold carrier
    _rMassLast : REAL := 0.0;          // 上次有效质量 [kg] / Last valid mass
    _rMassPrv  : REAL;                 // 上拍质量 [kg]（反流判据基准）/ Previous mass for backflow test
    _rTareInt  : REAL := 0.0;          // 皮重内部量 [kg] / Internal tare register
    _rFilled   : REAL;                 // 已注液量中间量 [kg] / Filled mass working value
    _rRemain   : REAL;                 // 剩余量中间量 [kg] / Remaining mass working value
    _rDriftRef : REAL;                 // 静置起始质量参照 [kg] / Dwell-start mass reference
    _bNearTgt  : BOOL;                 // 预关带迟滞判据回传保持变量 / Hysteresis pre-close band hold member
    _bMassBad  : BOOL;                 // 质量非有限标志 / Mass non-finite flag
    _uFault    : UDINT;                // 故障码锁存 / Latched fault code
    _uInfo     : UDINT;                // 信息码，每拍重算 / Info code
    _bFault    : BOOL;                 // 故障锁存位 / Latched fault bit
    _bCfgBad   : BOOL;                 // 组态非法聚合 / Configuration invalid aggregate
END_VAR
VAR CONSTANT
    DL_EF_INF_CAP  : REAL := 1.0E15;  // 非有限值筛查幅值上限 / Non-finite screening cap
    DL_EF_VALVE_OPEN  : REAL := 100.0;  // 粗注阀开度 [%] / Bulk fill valve opening
    DL_EF_VALVE_TRIM  : REAL := 30.0;   // 微调阀开度 [%] / Trim valve opening
END_VAR

(* —— 段 0：定时器与边沿实例无条件周期刷新（R182：调用语句不得置于 IF/CASE 内） —— *)
rtStart(CLK := bStart);                                                 // 启动沿刷新，每拍必调
rtReset(CLK := bReset);                                                 // 复位沿刷新，每拍必调
tonTareTo(IN := (_eState = E_DL_ElytFillState.eTare), PT := tTareTo);       // 皮重超时（单相独占）
tonFillTo(IN := (_eState = E_DL_ElytFillState.eFill), PT := tFillTo);       // 粗注超时（单相独占）
tonTrimTo(IN := (_eState = E_DL_ElytFillState.eTrim), PT := tTrimTo);       // 微调超时（单相独占）
tonDwell(IN := (_eState = E_DL_ElytFillState.eDwell), PT := tDwellTime);    // 浸润计时（单相独占，PT=配方时长）

(* —— 段 1：单拍量预清零（锁存量 _uFault/_bFault/_rTareInt/_rDriftRef 不入清单，R187①） —— *)
_uInfo := 16#0000_0000;             // 信息码每拍重算
bFillDone := FALSE;                 // 完成出口缺省 FALSE（Done 相单点置位）
bDwellDone := FALSE;                // 静置完成出口缺省 FALSE（Done 相单点置位）
_bCfgBad := FALSE;                  // 组态非法预清零
nErrId := 16#0000_0000;             // 事件码缺省无事件

(* —— 段 2：组态域闸（覆盖全部参与判据换算的引脚，R151） —— *)
IF (fBatchTargetKg <> fBatchTargetKg) OR (fBatchTargetKg <= 0.0) OR (ABS(fBatchTargetKg) > DL_EF_INF_CAP)
   OR (fFillTolKg <= 0.0) OR (fPrefillKg <= 0.0) OR (fHystKg <= 0.0)
   OR (fStatTolKg <= 0.0) OR (fDwellDriftKg <= 0.0)
   OR (TIME_TO_DINT(tTareTo) <= 0) OR (TIME_TO_DINT(tFillTo) <= 0)
   OR (TIME_TO_DINT(tTrimTo) <= 0) OR (TIME_TO_DINT(tDwellTime) <= 0) THEN
    _bCfgBad := TRUE;               // 目标/容差/提前量/漂移阈/时长域非法
END_IF

(* —— 段 3：eFault 迁出沿（R228-B：rtReset.Q 为输入引脚，恒可达） —— *)
IF rtReset.Q THEN
    _bFault := FALSE;               // 清故障锁存位
    _uFault := 16#0000_0000;
    IF _eState = E_DL_ElytFillState.eFault THEN
        _eState := E_DL_ElytFillState.eIdle;    // 故障相迁出：回空闲
    END_IF
END_IF

(* —— 段 4：质量采集与减量法换算（非有限保持；反流判据） —— *)
_bMassBad := (fTankMassKg <> fTankMassKg) OR (ABS(fTankMassKg) > DL_EF_INF_CAP) OR ((fTankMassKg - fTankMassKg) <> 0.0);
IF _bMassBad THEN
    _rMassEff := _rMassLast;        // 非有限：保持上次有效值
ELSE
    _rMassEff := fTankMassKg;       // 有效值入载体
    _rMassLast := fTankMassKg;
END_IF
IF (NOT _bMassBad) AND (_rMassEff - _rMassPrv > fStatTolKg) AND (_eState = E_DL_ElytFillState.eFill) THEN
    _uFault := 16#0006_04B7;        // 故障级：注液期质量上升（反流）
    _bFault := TRUE;
END_IF
_rMassPrv := _rMassEff;             // 反流判据基准更新（段尾单点）
IF NOT _bMassBad THEN
    _rFilled := _rTareInt - _rMassEff;          // 减量法：注液量 = 皮重 − 实时质量
ELSE
    _rFilled := 0.0;                // 质量无效：注液量出口置 0（防御口径）
END_IF
_rRemain := fBatchTargetKg - _rFilled;          // 剩余量
fFilledKg := _rFilled;              // 注液量出口镜像
fRemainingKg := _rRemain;           // 剩余量出口镜像
fTareKg := _rTareInt;               // 皮重出口镜像

(* —— 段 5：依赖件无条件周期刷新（容差窗 + 稳定窗 + 迟滞判据） —— *)
fbTol(bEnable := (_eState = E_DL_ElytFillState.eTrim),      // 仅微调相判定
      fTarget := fBatchTargetKg,                            // 目标注液量
      fActual := _rFilled,                                  // 实际注液量
      fTolerance := fFillTolKg,                             // 容差半宽
      fHysteresis := fHystKg);                              // 迟滞带（出窗防抖）
fbStat(fIn := _rMassEff,                                    // 质量稳定统计窗
       bSample := (_eState = E_DL_ElytFillState.eTare) OR (_eState = E_DL_ElytFillState.eDwell),
       nWindow := 32,                                       // 窗长（稳定判据标准口径）
       bClear := rtStart.Q);                                // 启动沿清窗（新批次重开）
_bNearTgt := FC_DL_Hysteresis(fIn := -_rRemain,             // 取反口径：剩余量落入预关带为 TRUE
                              fThreshold := -fPrefillKg,    // 预关阈（取反）
                              fHysteresis := fHystKg,       // 迟滞带（负值取绝对值语义由件内防御）
                              bState := _bNearTgt);         // 回传保持变量（同一成员，有状态纪律）

(* —— 段 6：相位机（只做迁移与阀指令；出口在段 8） —— *)
CASE _eState OF

E_DL_ElytFillState.eIdle:
    rValveCmdPct := 0.0;                    // 空闲：阀全关
    IF rtStart.Q AND _bCfgBad THEN
        _uFault := 16#0006_02B7;            // 故障级：组态非法
        _bFault := TRUE;
        _eState := E_DL_ElytFillState.eFault;
    ELSIF rtStart.Q AND (NOT _bCfgBad) THEN
        _rDriftRef := 0.0;                  // 静置参照预清零
        _eState := E_DL_ElytFillState.eTare;    // 进皮重相
    END_IF

E_DL_ElytFillState.eTare:
    rValveCmdPct := 0.0;                    // 皮重相：阀全关
    IF NOT _bMassBad THEN
        IF fbStat.bValid AND (fbStat.fRange <= fStatTolKg) THEN
            _rTareInt := _rMassEff;         // 锁皮重（稳定峰峰在阈内）
            _eState := E_DL_ElytFillState.eFill;    // 进粗注相
        ELSE
            _uInfo := 16#0006_07B7;         // 信息级：皮重稳定判据等待中
        END_IF
    END_IF
    IF tonTareTo.Q AND (_eState = E_DL_ElytFillState.eTare) THEN
        _uFault := 16#0006_03B7;            // 故障级：皮重相超时
        _bFault := TRUE;
        _eState := E_DL_ElytFillState.eFault;
    END_IF

E_DL_ElytFillState.eFill:
    rValveCmdPct := DL_EF_VALVE_OPEN;       // 粗注：阀全开
    IF tonFillTo.Q THEN
        _uFault := 16#0006_03B7;            // 故障级：粗注相超时
        _bFault := TRUE;
        rValveCmdPct := 0.0;                // 安全侧关阀
        _eState := E_DL_ElytFillState.eFault;
    ELSIF _bNearTgt THEN
        _eState := E_DL_ElytFillState.eTrim;    // 剩余量入预关带：进微调相
    END_IF

E_DL_ElytFillState.eTrim:
    IF _rRemain > 0.0 THEN
        rValveCmdPct := DL_EF_VALVE_TRIM;   // 微调：小开度收口
    ELSE
        rValveCmdPct := 0.0;                // 越量：关阀
    END_IF
    IF fbTol.bOk THEN
        rValveCmdPct := 0.0;                // 入容差带：关阀
        _rDriftRef := _rMassEff;            // 静置起始质量参照锁定
        _eState := E_DL_ElytFillState.eDwell;   // 进静置相
    ELSIF tonTrimTo.Q THEN
        _uFault := 16#0006_03B7;            // 故障级：微调相超时
        _bFault := TRUE;
        rValveCmdPct := 0.0;                // 安全侧关阀
        _eState := E_DL_ElytFillState.eFault;
    END_IF

E_DL_ElytFillState.eDwell:
    rValveCmdPct := 0.0;                    // 静置：阀全关
    IF ABS(_rMassEff - _rDriftRef) > fDwellDriftKg THEN
        _uInfo := 16#0006_06B7;             // 信息级：静置漂移超阈（渗漏提示，不置故障）
    END_IF
    IF tonDwell.Q THEN
        _eState := E_DL_ElytFillState.eDone;    // 浸润到点：进完成相
    END_IF

E_DL_ElytFillState.eDone:
    rValveCmdPct := 0.0;                    // 完成：阀全关
    bFillDone := TRUE;                      // 完成出口（Done 相每拍重申）
    bDwellDone := TRUE;                     // 静置完成出口（Done 相每拍重申）
    _uInfo := 16#0006_01B7;                 // 信息级：周期完成
    IF NOT bStart THEN
        _eState := E_DL_ElytFillState.eIdle;    // 指令撤销：回空闲
    END_IF

E_DL_ElytFillState.eFault:
    rValveCmdPct := 0.0;                    // 故障相：阀全关（安全侧）
    ;                                       // 等复位沿（段 3 承载迁出）

ELSE
    _uFault := 16#0006_05B7;                // 故障级：非法相位 ID 兜底
    _bFault := TRUE;
    rValveCmdPct := 0.0;                    // 安全侧关阀
    _eState := E_DL_ElytFillState.eFault;   // 强制回故障相

END_CASE

(* —— 段 7：称重非有限持续判故障（段 4 标志的锁存化，R228-B 配对） —— *)
IF _bMassBad AND (_eState <> E_DL_ElytFillState.eIdle) THEN
    _uFault := 16#0006_04B7;                // 故障级：称重信号非有效持续（活动相内）
    _bFault := TRUE;
END_IF

(* —— 段 8：出口单点映射（名实同源；锁存码回放，禁同拍抹除） —— *)
IF _bFault THEN
    nErrId := _uFault;                      // 故障锁存码回放（不在故障相按当下输入重推）
    bFillDone := FALSE;                     // 故障相完成出口强制 FALSE（安全侧）
    bDwellDone := FALSE;
ELSE
    nErrId := _uInfo;                       // 信息码
END_IF
eState := _eState;                          // 状态出口单点映射

END_FUNCTION_BLOCK

(* ---- FB_DL_ElectrolyteFillVacuum.st ---- *)
(*==============================================================================
 * 组件名称 (Component)  : FB_DL_ElectrolyteFillVacuum
 * 所属子库 (Sublibrary) : DL_Process
 * 当前版本 (Version)    : 1.0.0
 * 兼容性 (Platform)     : CODESYS 3.5+ / TwinCAT 3 / 汇川 InoProShop / 施耐德 Machine Expert
 *                         仅依赖 Standard.library（TON / R_TRIG / ABS），零厂商私有库
 * 功能描述 (Function)   : 注液真空度监视与静置计时台账。注液运行电平内监视
 *                         真空度对设定容差窗（bVacOk），静置 TON 达 tHoldReq
 *                         即 bHoldDone；静置期记录最低真空度台账；注液结束
 *                         沿若静置已完成则批次计数 +1 并清窗内台账。与
 *                         VacuumGaugeMux（计融合）分工：本件是静置窗 + 门限
 *                         + 批次计数的工艺台账件。
 * 来源标签 (Origin)     : ROADMAP §21.1 R13 池（L879），自研 clean-room
 * 边界语义 (Boundary)   : ① 真空度 NaN/Inf 拍：bVacOk 强制 FALSE（安全侧，
 *                         静置计时断链不误完成）；
 *                         ② 容差/静置时长/秒值域闸 → 组态故障；
 *                         ③ 最低真空台账随静置起步清零、随批次收口清零；
 *                         ④ TON 为电平计时（非自复位周期窗）。
 * 输出语义 (Fallback)   : 【R191】bEnable = FALSE → bVacOk/bHoldDone 强制
 *                         FALSE（监视出口失能必须收敛）；eFault 相 → FALSE
 *                         + bError = TRUE。
 * 码位     (Codes)      : 按 R297 范式零 16# 码位硬编码；错误出口 BOOL+ENUM(eCause)。
 * 红线自检 (Redline)    : 7 项红线已自检：R1 零全局 ✓｜R2 零物理地址 ✓｜R3 纯 IEC ✓
 *                         R4 除零无涉/NaN 安全侧/组态闸 ✓｜R5 双语同行注释 ✓
 *                         R6 CASE 带 ELSE 兜底迁 eFault ✓｜R7 TON/R_TRIG 段 0 无条件刷新 ✓
 * 验收向量 (Acceptance) : V1 设定 5.0 kPa 容差 0.5、实测 5.2 → bVacOk=TRUE，
 *                         静置 T#60S 到时 → bHoldDone=TRUE；
 *                         V2 静置期实测最低 4.3 → fVacMinHold=4.3；
 *                         V3 bFillEnd 沿且静置已完成 → nBatchCnt+1 且台账清零。
 * 修订历史 (Revision)   : 2026-11-20  v1.0.0  R51 首版（批 3 · 序号 12）
 *==============================================================================*)
TYPE E_DL_EfvState :
(
    eIdle  := 0,                             (* 待使能 / Idle *)
    eFill  := 10,                            (* 注液监视运行 / Fill monitor *)
    eFault := 90                             (* 故障锁存相 / Fault latched phase *)
);
END_TYPE

TYPE E_DL_EfvCause :
(
    eNone       := 0,                        (* 无故障成因 / No cause *)
    eCfgIllegal := 1,                        (* 组态非法：容差/时长/秒值越域 / Illegal config *)
    ePhaseBad   := 2                         (* 非法相位兜底 / Illegal phase fallback *)
);
END_TYPE

FUNCTION_BLOCK FB_DL_ElectrolyteFillVacuum
VAR_INPUT
    fVacKpa   : LREAL := 0.0;                (* 真空度实测 [kPa] / Vacuum actual *)
    fVacSp    : LREAL := 5.0;                (* 真空度设定 [kPa] / Vacuum setpoint *)
    fVacTol   : LREAL := 0.5;                (* 真空容差，域 > 0 [kPa] / Vacuum tolerance *)
    tHoldReq  : TIME := T#60S;               (* 静置时长要求，域 > T#0S [ms] / Hold time requirement *)
    bFillRun  : BOOL := FALSE;               (* 注液运行电平 [-] / Fill run level *)
    bFillEnd  : BOOL := FALSE;               (* 注液结束沿 [-] / Fill end edge *)
    bEnable   : BOOL := TRUE;                (* 使能 [-] / Enable *)
    bReset    : BOOL := FALSE;               (* 复位命令，上升沿清全部 [-] / Reset command *)
END_VAR
VAR_OUTPUT
    bVacOk    : BOOL;                        (* 真空度在容差窗内 [-] / Vacuum in tolerance *)
    bHoldDone : BOOL;                        (* 静置完成（TON 到时电平）[-] / Hold done *)
    fVacMinHold: LREAL;                      (* 本次静置期最低真空度台账 [kPa] / Min vacuum ledger *)
    tHoldElapsed : TIME;                     (* 静置已进行时长（诊断）[ms] / Hold elapsed *)
    nBatchCnt : UDINT;                       (* 完成批次计数（静置完 + 结束沿）[批] / Batch count *)
    eState    : E_DL_EfvState;               (* 状态出口 / State outlet *)
    eCause    : E_DL_EfvCause;               (* 故障成因出口 / Fault cause outlet *)
    bError    : BOOL;                        (* 故障锁存标志 [-] / Fault latch flag *)
END_VAR
VAR
    _eState   : E_DL_EfvState := E_DL_EfvState.eIdle;     (* 内部相位（CASE 唯一写入目标） / Internal phase *)
    _eCause   : E_DL_EfvCause := E_DL_EfvCause.eNone;     (* 故障成因锁存量 / Latched cause *)
    rtEnd     : R_TRIG;                      (* 结束沿实例，段 0 无条件调用 / End edge instance *)
    rtReset   : R_TRIG;                      (* 复位沿实例，段 0 无条件调用 / Reset edge instance *)
    tonHold   : TON;                         (* 静置计时，段 0 无条件调用 / Hold timer *)
    _fVacMin  : LREAL;                       (* 最低真空锁存 [kPa] / Min vacuum latch *)
    _bHoldL   : BOOL;                        (* 静置完成锁存（结转批次判据）[-] / Hold-done latch *)
    _nBatch   : UDINT;                       (* 批次计数锁存 [批] / Batch count latch *)
    _bVacBad  : BOOL;                        (* 真空非有限当拍量 [-] / Non-finite vacuum *)
    _bFault   : BOOL;                        (* 故障锁存位 / Latched fault bit *)
    _bCfgBad  : BOOL;                        (* 组态非法当拍量 / Illegal config this scan *)
END_VAR
VAR CONSTANT
    DL_EFV_EPS : LREAL := 1.0E-9;            (* 容差判零容差 [kPa] / Tolerance epsilon *)
END_VAR

(* —— 段 0：当拍判据派生 + 实例无条件刷新（R228A） —— *)
_bCfgBad := (fVacTol <= DL_EFV_EPS) OR (tHoldReq <= T#0S);   (* 组态闸（R151 全引脚） / Config gate *)
rtEnd(CLK := bFillEnd);                      (* 结束沿每拍必调 / End edge every scan *)
rtReset(CLK := bReset);                      (* 复位沿每拍必调 / Reset edge every scan *)
_bVacBad := (fVacKpa <> fVacKpa) OR ((fVacKpa - fVacKpa) <> (fVacKpa - fVacKpa));   (* 真空 NaN 自反 + Inf 差判 / Non-finite vacuum *)
tonHold(IN := (_eState = E_DL_EfvState.eFill) AND bFillRun AND (NOT _bVacBad) AND bVacOk, PT := tHoldReq);   (* 静置计时：容差窗内才走时（电平计时非周期窗） / Hold timer, gated by window *)

(* —— 段 1：单拍量预清零（R107） —— *)
bVacOk := FALSE;                             (* 真空判定预清（全路径赋值） / Vac-ok preset *)
bHoldDone := FALSE;                          (* 静置完成预清 / Hold-done preset *)

(* —— 段 2：复位沿处理（作用域：清故障 + 清批次计数 + 清台账 + 清锁存 + 迁 eIdle，R283 逐项声明） —— *)
IF rtReset.Q THEN
    _bFault := FALSE;                        (* 清故障锁存 / Clear fault *)
    _eCause := E_DL_EfvCause.eNone;          (* 清成因 / Clear cause *)
    _nBatch := 0;                            (* 清批次计数 / Clear batch count *)
    _fVacMin := 0.0;                         (* 清最低台账 / Clear min ledger *)
    fVacMinHold := 0.0;                      (* 清台账出口 / Clear ledger outlet *)
    _bHoldL := FALSE;                        (* 清静置锁存 / Clear hold latch *)
    _eState := E_DL_EfvState.eIdle;          (* 迁待机相 / Back to idle *)
END_IF

(* —— 段 3：组态闸故障锁存（R45 配对；锁存至复位沿，R189） —— *)
IF _bCfgBad AND NOT _bFault THEN
    _bFault := TRUE;                         (* 锁存故障位 / Latch fault *)
    _eCause := E_DL_EfvCause.eCfgIllegal;    (* 成因：组态非法 / Cause: illegal config *)
    _eState := E_DL_EfvState.eFault;         (* 同步迁故障相 / Migrate to fault *)
END_IF

(* —— 段 4：CASE 主状态机（ELSE 兜底迁 eFault，红线 6） —— *)
CASE _eState OF
    E_DL_EfvState.eIdle:                     (* 待机相 / Idle *)
        IF bEnable AND NOT _bFault THEN
            _eState := E_DL_EfvState.eFill;  (* 进入监视 / Enter fill *)
        END_IF
    E_DL_EfvState.eFill:                     (* 监视相：容差判定 + 静置 + 台账 + 批次收口 / Fill *)
        IF NOT bEnable THEN
            _eState := E_DL_EfvState.eIdle;  (* 失能回待机 / Back to idle *)
        ELSE
            IF NOT _bVacBad THEN
                bVacOk := ABS(fVacKpa - fVacSp) <= fVacTol;   (* 容差窗判定（除法无涉） / Tolerance verdict *)
            END_IF                           (* 坏值拍 bVacOk 保持预清 FALSE（边界①安全侧） / Bad scan: safe FALSE *)
            bHoldDone := tonHold.Q;          (* 静置完成出口 / Hold-done outlet *)
            IF tonHold.Q AND (NOT _bHoldL) THEN   (* 静置完成沿：锁定 + 台账起步 / On hold-done edge *)
                _bHoldL := TRUE;             (* 置完成锁存（供批次收口结转） / Set hold latch *)
            END_IF
            IF bFillRun AND (NOT _bVacBad) AND bVacOk THEN   (* 静置期最低真空台账 / Min ledger *)
                IF (_fVacMin = 0.0) OR (fVacKpa < _fVacMin) THEN   (* 首样本或更低取值（0.0 为哨兵起点非合法真空读数） / First-or-lower *)
                    _fVacMin := fVacKpa;     (* 更新最低 / Update min *)
                END_IF
            END_IF
            IF rtEnd.Q THEN                  (* 注液结束沿：批次收口判定 / On fill end edge *)
                IF _bHoldL THEN
                    _nBatch := _nBatch + 1;  (* 静置已完成：批次 +1（UDINT 回绕工程安全） / Count batch *)
                    _bHoldL := FALSE;        (* 清完成锁存（下一批重新静置） / Clear hold latch *)
                END_IF
                _fVacMin := 0.0;             (* 清窗内台账（边界③：随收口清零） / Clear ledger *)
                fVacMinHold := _fVacMin;     (* 台账出口刷新 / Ledger outlet *)
            ELSE
                fVacMinHold := _fVacMin;     (* 台账出口实时镜像 / Ledger mirror *)
            END_IF
        END_IF
    E_DL_EfvState.eFault:                    (* 故障相：冻结保持，仅复位沿出 / Fault *)
        ;                                    (* 锁存回放（R28） / Replay from latch *)
    ELSE                                     (* 非法相位兜底迁安全态 / Illegal phase fallback *)
        _eState := E_DL_EfvState.eFault;     (* 迁故障相 / To fault *)
        _bFault := TRUE;                     (* 同步锁存 / Latch *)
        _eCause := E_DL_EfvCause.ePhaseBad;  (* 成因：非法相位 / Cause: illegal phase *)
END_CASE

(* —— 段 5：出口映射（bError/eState 同源，R191） —— *)
tHoldElapsed := tonHold.ET;                  (* 静置时长诊断镜像 / Elapsed mirror *)
nBatchCnt := _nBatch;                        (* 批次计数出口 / Batch outlet *)
bError := _bFault;                           (* 故障标志镜像 / Fault flag mirror *)
eState := _eState;                           (* 状态出口 / State outlet *)
eCause := _eCause;                           (* 成因出口 / Cause outlet *)
END_FUNCTION_BLOCK
